(* IEC 61131-3 sources: daoli-st-library/DL_Process (part 11) *)

(* ---- FC_DL_CompressorDutyCycleCalc.st ---- *)
(*
  ============================================================
  组件名 : FC_DL_CompressorDutyCycleCalc
  分类   : DL_Process
  功能   : 压缩机加载占空比与卸载能耗占比计算，用于评估空压站运行经济性
  复杂度 : C1
  版本   : 1.0.0
  作者   : 道莅工业代码库工厂 / R81
  日期   : 2026-11-24
  开源溯源 : clean-room（no upstream）—— 依据公开工程公式自研，未复制任何上游实现
  红线自检 : R1 无GVL/R2 无物理地址/R3 纯IEC/R4 防除零/R5 双语注释
  接口说明 :
      加载占空比 = 加载时间 / 统计窗口 * 100。
      卸载能耗占比 = 卸载功率*卸载时间 / (加载功率*加载时间 + 卸载功率*卸载时间) * 100。
      能耗分母为零表示窗口内既无加载也无卸载，占空比无法归一，判无效。
      加载时间加卸载时间超过统计窗口时数据自相矛盾，判无效而不是强行归一。
  ============================================================
*)
FUNCTION FC_DL_CompressorDutyCycleCalc : BOOL
VAR_INPUT
    bEnable      : BOOL; // 使能：TRUE 时计算 / Enable: TRUE to compute
    bErr         : BOOL; // 外部故障：TRUE 时立即退出并置结果无效 / External fault: TRUE aborts with invalid result
    rLoadTime_s  : REAL; // 窗口内加载运行时间 [s] / loaded running time inside the window [second]
    rUnloadTime_s : REAL; // 窗口内卸载运行时间 [s] / unloaded running time inside the window [second]
    rIdleKw      : REAL; // 卸载空转功率 [kW] / unloaded idle power [kilowatt]
    rLoadKw      : REAL; // 加载运行功率 [kW] / loaded running power [kilowatt]
    rDur_s       : REAL; // 统计窗口总时长 [s] / total duration of the statistic window [second]
END_VAR
VAR_OUTPUT
    rDutyPct       : REAL; // 加载占空比，限幅 0~100 [%] / loading duty cycle clamped to 0 to 100 [percent]
    rIdleEnergyPct : REAL; // 卸载能耗占窗口总能耗比例，限幅 0~100 [%] / unloaded energy share of the window total clamped to 0 to 100 [percent]
    rTotalKwh      : REAL; // 窗口内折算总电量 [kWh] / equivalent total energy inside the window [kilowatt hour]
    bValid         : BOOL; // 输出有效：TRUE 表示结果可用 / Output valid
END_VAR
VAR CONSTANT
    DL_R_MAX   : REAL := 3.0E38;  // 实数上界，用于拦截 Inf [无量纲] / real upper bound used to reject infinity [dimensionless]
    DL_EPS     : REAL := 1.0E-12; // 除零判定阈值 [无量纲] / division guard threshold [dimensionless]
    DL_PCT     : REAL := 100.0;   // 百分数换算系数 [无量纲] / percentage scaling factor [dimensionless]
    DL_ZERO    : REAL := 0.0;     // 零值常量 [无量纲] / zero constant [dimensionless]
    DL_S_PER_H : REAL := 3600.0;  // 每小时秒数 [s/h] / seconds per hour [second per hour]
    DL_TOL_S   : REAL := 0.001;   // 时间窗超限判定容差 [s] / tolerance for the window overrun check [second]
END_VAR
VAR
    _bFin    : BOOL := FALSE; // 输入有限性判定结果 / input finiteness verdict
    _rLoadKwh : REAL := 0.0;  // 加载段电量 [kWh] / energy of the loaded segment [kilowatt hour]
    _rIdleKwh : REAL := 0.0;  // 卸载段电量 [kWh] / energy of the unloaded segment [kilowatt hour]
    _rDen     : REAL := 0.0;  // 能耗占比分母 [kWh] / denominator of the energy share [kilowatt hour]
END_VAR

    // 段 1｜出口预置
    rDutyPct := 0.0;
    rIdleEnergyPct := 0.0;
    rTotalKwh := 0.0;
    bValid := FALSE;
    // 段 2｜使能闸与外部故障闸
    IF NOT bEnable THEN
        RETURN;
    END_IF;
    IF bErr THEN
        RETURN;
    END_IF;
    // 段 3｜非有限闸
    _bFin := (rLoadTime_s = rLoadTime_s) AND (ABS(rLoadTime_s) <= DL_R_MAX) AND (rUnloadTime_s = rUnloadTime_s) AND (ABS(rUnloadTime_s) <= DL_R_MAX) AND (rIdleKw = rIdleKw) AND (ABS(rIdleKw) <= DL_R_MAX) AND (rLoadKw = rLoadKw) AND (ABS(rLoadKw) <= DL_R_MAX) AND (rDur_s = rDur_s) AND (ABS(rDur_s) <= DL_R_MAX);
    IF NOT _bFin THEN
        RETURN;
    END_IF;
    // 段 4｜域闸：统计窗口严格为正，时间与功率不得为负
    IF (ABS(rDur_s) <= DL_EPS) OR (rDur_s < DL_ZERO) THEN
        RETURN;
    END_IF;
    IF (rLoadTime_s < DL_ZERO) OR (rUnloadTime_s < DL_ZERO) OR (rIdleKw < DL_ZERO) OR (rLoadKw < DL_ZERO) THEN
        RETURN;
    END_IF;
    // 段 5｜加载加卸载不得超过窗口，超出部分属数据矛盾
    IF (rLoadTime_s + rUnloadTime_s) > (rDur_s + DL_TOL_S) THEN
        RETURN;
    END_IF;
    // 段 6｜加载占空比与限幅
    rDutyPct := rLoadTime_s / rDur_s * DL_PCT;
    IF rDutyPct < DL_ZERO THEN
        rDutyPct := DL_ZERO;
    END_IF;
    IF rDutyPct > DL_PCT THEN
        rDutyPct := DL_PCT;
    END_IF;
    // 段 7｜两段电量与总电量
    _rLoadKwh := rLoadKw * rLoadTime_s / DL_S_PER_H;
    _rIdleKwh := rIdleKw * rUnloadTime_s / DL_S_PER_H;
    rTotalKwh := _rLoadKwh + _rIdleKwh;
    // 段 8｜能耗占比分母闸
    _rDen := _rLoadKwh + _rIdleKwh;
    IF _rDen <= DL_EPS THEN
        RETURN;
    END_IF;
    rIdleEnergyPct := _rIdleKwh / _rDen * DL_PCT;
    IF rIdleEnergyPct < DL_ZERO THEN
        rIdleEnergyPct := DL_ZERO;
    END_IF;
    IF rIdleEnergyPct > DL_PCT THEN
        rIdleEnergyPct := DL_PCT;
    END_IF;
    bValid := TRUE;
    FC_DL_CompressorDutyCycleCalc := bValid;
END_FUNCTION

(* ---- FC_DL_ConductivityDilutionCalc.st ---- *)
(*
  ============================================================
  组件名 : FC_DL_ConductivityDilutionCalc
  分类   : DL_Process
  功能   : 电导率稀释比计算，由母液与水的本底电导求目标浓度所需的稀释倍数与配水占比
  复杂度 : C1
  版本   : 1.0.0
  作者   : 道莅工业代码库工厂 / R81
  日期   : 2026-11-24
  开源溯源 : clean-room（no upstream）—— 依据公开工程公式自研，未复制任何上游实现
  红线自检 : R1 无GVL/R2 无物理地址/R3 纯IEC/R4 防除零/R5 双语注释
  接口说明 :
      稀释比 = (母液电导 - 水本底电导) / (目标电导 - 水本底电导)。
      目标电导不高于水本底时分母非正，物理上无法靠兑水达到，直接判无效。
      配水占比 = (1 - 1/稀释比) * 100，稀释比非正时同样判无效。
  ============================================================
*)
FUNCTION FC_DL_ConductivityDilutionCalc : BOOL
VAR_INPUT
    bEnable      : BOOL; // 使能：TRUE 时计算 / Enable: TRUE to compute
    bErr         : BOOL; // 外部故障：TRUE 时立即退出并置结果无效 / External fault: TRUE aborts with invalid result
    rCondFeed    : REAL; // 母液电导率 [uS/cm] / feed solution conductivity [micro siemens per centimetre]
    rCondTarget  : REAL; // 目标电导率 [uS/cm] / target conductivity [micro siemens per centimetre]
    rCondWater   : REAL; // 稀释水本底电导率 [uS/cm] / background conductivity of the dilution water [micro siemens per centimetre]
END_VAR
VAR_OUTPUT
    rDilutionRatio : REAL; // 稀释倍数，母液体积的多少倍 [无量纲] / dilution ratio in multiples of the feed volume [dimensionless]
    rWaterPct      : REAL; // 配水中水所占体积百分比 [%] / volumetric percentage of water in the mixture [percent]
    bValid         : BOOL; // 输出有效：TRUE 表示结果可用 / Output valid
END_VAR
VAR CONSTANT
    DL_R_MAX : REAL := 3.0E38;  // 实数上界，用于拦截 Inf [无量纲] / real upper bound used to reject infinity [dimensionless]
    DL_EPS   : REAL := 1.0E-12; // 除零判定阈值 [无量纲] / division guard threshold [dimensionless]
    DL_ONE   : REAL := 1.0;     // 单位常量 [无量纲] / unity constant [dimensionless]
    DL_PCT   : REAL := 100.0;   // 百分数换算系数 [无量纲] / percentage scaling factor [dimensionless]
    DL_RATIO_MAX : REAL := 10000.0; // 稀释比合理上限，超限视为配比不可实现 [无量纲] / sanity upper bound of the dilution ratio [dimensionless]
END_VAR
VAR
    _bFin  : BOOL := FALSE; // 输入有限性判定结果 / input finiteness verdict
    _rNum  : REAL := 0.0;   // 稀释比分子 [uS/cm] / numerator of the dilution ratio [micro siemens per centimetre]
    _rDen  : REAL := 0.0;   // 稀释比分母 [uS/cm] / denominator of the dilution ratio [micro siemens per centimetre]
END_VAR

    // 段 1｜出口预置
    rDilutionRatio := 0.0;
    rWaterPct := 0.0;
    bValid := FALSE;
    // 段 2｜使能闸与外部故障闸
    IF NOT bEnable THEN
        RETURN;
    END_IF;
    IF bErr THEN
        RETURN;
    END_IF;
    // 段 3｜非有限闸
    _bFin := (rCondFeed = rCondFeed) AND (ABS(rCondFeed) <= DL_R_MAX) AND (rCondTarget = rCondTarget) AND (ABS(rCondTarget) <= DL_R_MAX) AND (rCondWater = rCondWater) AND (ABS(rCondWater) <= DL_R_MAX);
    IF NOT _bFin THEN
        RETURN;
    END_IF;
    // 段 4｜域闸：三者均不得为负，母液必须高于水本底
    IF (rCondFeed < 0.0) OR (rCondTarget < 0.0) OR (rCondWater < 0.0) THEN
        RETURN;
    END_IF;
    // 段 5｜分子分母组装
    _rNum := rCondFeed - rCondWater;
    _rDen := rCondTarget - rCondWater;
    // 段 6｜分母非正闸：兑水无法把电导降到水本底以下
    IF _rDen <= DL_EPS THEN
        RETURN;
    END_IF;
    // 段 7｜分子非正闸：母液不高于水本底时无稀释意义
    IF _rNum <= DL_EPS THEN
        RETURN;
    END_IF;
    rDilutionRatio := _rNum / _rDen;
    // 段 8｜稀释比合理区间闸，防止配比不可实现
    IF (rDilutionRatio < DL_ONE) OR (rDilutionRatio > DL_RATIO_MAX) THEN
        RETURN;
    END_IF;
    // 段 9｜配水占比
    rWaterPct := (DL_ONE - DL_ONE / rDilutionRatio) * DL_PCT;
    IF rWaterPct < 0.0 THEN
        rWaterPct := 0.0;
    END_IF;
    IF rWaterPct > DL_PCT THEN
        rWaterPct := DL_PCT;
    END_IF;
    bValid := TRUE;
    FC_DL_ConductivityDilutionCalc := bValid;
END_FUNCTION

(* ---- FC_DL_CoreSandBakeCurveCalc.st ---- *)
(*
 * FC_DL_CoreSandBakeCurveCalc | C2 | DL_Process
 * 功能：芯砂烘干升温曲线（升温段、总时间）与保温后残余水分       单位：温度 [℃]、升温速率 [K/min]、时间 [min]、水分 [%]
 * 工况边界：升温段按线性斜坡、保温段按一阶指数衰减残余水分 res=1.5×EXP(−hold/40)；升温速率须 >0、目标温度须高于起始温度，否则判 9716；本件不含分段升温与露点控制
 * 代数值回代：target=200、start=25、rate=3 → ramp=175/3=58.33 min；total=58.33+60=118.33 min；res=1.5×EXP(−60/40)=1.5×0.2231=0.335 %（spec 记 0.33 %，一致）
 * 开源溯源：clean-room 自研，未复制任何第三方代码（无外部来源）
 *)
FUNCTION FC_DL_CoreSandBakeCurveCalc : BOOL
VAR_INPUT
    rTargetC   : REAL := 200.0;      // 目标烘干温度 | target baking temperature [℃]
    rRampKmin  : REAL := 3.0;        // 升温速率 | heating rate [K/min]
    rStartC    : REAL := 25.0;       // 起始温度 | starting temperature [℃]
    rHoldMin   : REAL := 60.0;       // 保温时间 | holding time [min]
END_VAR
VAR_OUTPUT
    rRampMin        : REAL;          // 升温段时间 | ramp duration [min]
    rTotalMin       : REAL;          // 总时间（升温+保温）| total time, ramp plus hold [min]
    rResidualMoistPct : REAL;        // 保温后残余水分 | residual moisture after holding [%]
    xValid          : BOOL;          // 输出有效 | outputs valid
    nFaultCode      : INT;           // 0=无 / 9716=温度或速率非法 | 0 none, 9716 illegal temperature or rate
END_VAR
VAR
    xFinTg  : BOOL;                  // 目标温度有限性 | target temperature is finite
    xFinRt  : BOOL;                  // 升温速率有限性 | heating rate is finite
    xFinSt  : BOOL;                  // 起始温度有限性 | starting temperature is finite
    xFinHd  : BOOL;                  // 保温时间有限性 | holding time is finite
END_VAR
VAR CONSTANT
    DL_CSB_MOIST0   : REAL := 1.5;   // 保温起始残余水分基准 | residual moisture at the start of holding [%]
    DL_CSB_TAU_MIN  : REAL := 40.0;  // 水分衰减时间常数 | moisture decay time constant [min]
END_VAR

// 段1｜非有限闸（R19）
xFinTg := (rTargetC = rTargetC) AND ((rTargetC - rTargetC) = 0.0);
xFinRt := (rRampKmin = rRampKmin) AND ((rRampKmin - rRampKmin) = 0.0);
xFinSt := (rStartC = rStartC) AND ((rStartC - rStartC) = 0.0);
xFinHd := (rHoldMin = rHoldMin) AND ((rHoldMin - rHoldMin) = 0.0);
IF (NOT xFinTg) OR (NOT xFinRt) OR (NOT xFinSt) OR (NOT xFinHd) THEN
    rRampMin := 0.0;                 // 安全值：时间 0 | safe value, zero times
    rTotalMin := 0.0;
    rResidualMoistPct := 0.0;
    xValid := FALSE;
    nFaultCode := 9716;
    FC_DL_CoreSandBakeCurveCalc := FALSE;
    RETURN;
END_IF

// 段2｜域闸：速率入分母须 >0，目标须高于起始，保温时间非负
IF (rRampKmin <= 0.0) OR (rTargetC <= rStartC) OR (rHoldMin < 0.0) THEN
    rRampMin := 0.0;
    rTotalMin := 0.0;
    rResidualMoistPct := 0.0;
    xValid := FALSE;
    nFaultCode := 9716;
    FC_DL_CoreSandBakeCurveCalc := FALSE;
    RETURN;
END_IF

// 段3｜算法：ramp=(target−start)/rate；total=ramp+hold；res=1.5×EXP(−hold/40)
rRampMin := (rTargetC - rStartC) / rRampKmin;
rTotalMin := rRampMin + rHoldMin;
rResidualMoistPct := DL_CSB_MOIST0 * EXP(-rHoldMin / DL_CSB_TAU_MIN);

// 段4｜出口
nFaultCode := 0;
xValid := TRUE;
FC_DL_CoreSandBakeCurveCalc := TRUE;
END_FUNCTION

(* ---- FC_DL_CrusherThroughputCalc.st ---- *)
(*
  Name: FC_DL_CrusherThroughputCalc
  Category: DL_Process
  Version: 1.0.0
  Round: R89 / 2026-11-25
  开源溯源：clean-room 自研（族 矿山破碎筛分，ST 开源生态实测 0 命中，无外部代码引入）
  功能：按排矿口开口比产能法算颚式/圆锥破碎机实际产能，并以单程合格率反算闭路循环负荷率。
  边界条件：① 五入参全部过非有限闸（NaN 自反判 / Inf 差值自减判），任一非有限返回哨兵 -1；
            ② 排矿口 < 3 mm 或给料粒度不高于排矿口 1.2 倍（无有效破碎比）判组态非法，返回哨兵 -1；
            ③ 单程合格率下限 0.1，循环负荷率钳位 0~500 %（钳的是量值不钳事实，有效性不受影响）。
  量纲自证：q0[t/(h·mm)] × gap[mm] = t/h；kH / kD 无量纲；CL=(1/p−1)×100 无量纲。
*)
FUNCTION FC_DL_CrusherThroughputCalc : REAL
VAR_INPUT
    fFeedTph : REAL;        (* 给料量（新给矿） [t/h] Feed rate, fresh feed *)
    fGapMm : REAL;          (* 排矿口开口（闭侧） [mm] Closed-side gap [mm] *)
    fFeedSizeMm : REAL;     (* 给料粒度（95% 通过粒径） [mm] Feed size, 95% passing *)
    fHardnessIdx : REAL;    (* 硬度指数（1.0 为基准矿） [-] Hardness index, 1.0 baseline *)
    fBulkDensity : REAL;    (* 堆密度 [t/m3] Bulk density [t/m3] *)
END_VAR
VAR_OUTPUT
    fThroughputTph : REAL;      (* 实际破碎通过量 [t/h] Actual throughput [t/h] *)
    fCirculatingLoadPct : REAL; (* 闭路循环负荷率 [%] Circulating load ratio [%] *)
    xValid : BOOL;              (* 计算有效性标志 [-] Calculation valid flag *)
END_VAR
VAR CONSTANT
    DL_EPS : REAL := 1.0E-9;        (* 除零判定容差 [-] Divide-by-zero tolerance *)
    DL_Q0 : REAL := 2.5;            (* 单位开口基准产能 [t/(h·mm)] Specific capacity per gap *)
    DL_DENS_REF : REAL := 1.6;      (* 基准堆密度 [t/m3] Reference bulk density *)
    DL_RR_MIN : REAL := 1.2;        (* 最小有效破碎比 [-] Minimum reduction ratio *)
    DL_CL_MAX : REAL := 500.0;      (* 循环负荷率饱和上限 [%] Circulating load ceiling *)
    DL_PASS_MIN : REAL := 0.1;      (* 单程合格率下限 [-] Minimum single-pass fraction *)
    DL_GAP_MIN : REAL := 3.0;       (* 排矿口工程下限 [mm] Minimum engineering gap *)
    DL_H_MIN : REAL := 0.2;         (* 硬度指数下限 [-] Hardness index floor *)
    DL_H_MAX : REAL := 5.0;         (* 硬度指数上限 [-] Hardness index ceiling *)
    DL_D_MIN : REAL := 0.5;         (* 堆密度下限 [t/m3] Bulk density floor *)
    DL_D_MAX : REAL := 4.0;         (* 堆密度上限 [t/m3] Bulk density ceiling *)
END_VAR
VAR
    fRr : REAL;     (* 破碎比 = 给料粒度/排矿口 [-] Reduction ratio *)
    fKh : REAL;     (* 硬度修正系数 [-] Hardness correction factor *)
    fKd : REAL;     (* 密度修正系数 [-] Density correction factor *)
    fQcap : REAL;   (* 排矿口通过能力 [t/h] Gap capability [t/h] *)
    fPass : REAL;   (* 单程合格率 [-] Single-pass pass fraction *)
    fQout : REAL;   (* 当拍通过量中间量 [t/h] Throughput scratch [t/h] *)
END_VAR
(* 出口预置：三出口统一预置安全值（R256） *)
fThroughputTph := 0.0; fCirculatingLoadPct := 0.0; xValid := FALSE;
(* 非有限闸：NaN 自反判 + Inf 差值自减判，五入参全枚举（R272） *)
IF (fFeedTph <> fFeedTph) OR ((fFeedTph - fFeedTph) <> 0.0)
   OR (fGapMm <> fGapMm) OR ((fGapMm - fGapMm) <> 0.0)
   OR (fFeedSizeMm <> fFeedSizeMm) OR ((fFeedSizeMm - fFeedSizeMm) <> 0.0)
   OR (fHardnessIdx <> fHardnessIdx) OR ((fHardnessIdx - fHardnessIdx) <> 0.0)
   OR (fBulkDensity <> fBulkDensity) OR ((fBulkDensity - fBulkDensity) <> 0.0) THEN
    FC_DL_CrusherThroughputCalc := -1.0;    (* 哨兵 -1：入参非有限 / Sentinel -1, non-finite input *)
    RETURN;
END_IF
(* 组态域闸：给料、开口、粒度、硬度、密度逐项定域（禁 NaN 判假即放行，全用正向不等号） *)
IF (fFeedTph <= DL_EPS) OR (fGapMm < DL_GAP_MIN)
   OR (fFeedSizeMm <= fGapMm * DL_RR_MIN)
   OR (fHardnessIdx < DL_H_MIN) OR (fHardnessIdx > DL_H_MAX)
   OR (fBulkDensity < DL_D_MIN) OR (fBulkDensity > DL_D_MAX) THEN
    FC_DL_CrusherThroughputCalc := -1.0;    (* 哨兵 -1：组态非法 / Sentinel -1, bad configuration *)
    RETURN;
END_IF
(* 破碎比：给料粒度 ÷ 排矿口，除子已过工程下限闸，量纲 mm/mm = 无量纲 *)
fRr := fFeedSizeMm / fGapMm;
(* 硬度修正：kH = 1/(0.6+0.4·H)，H = 1.0 时恰为 1.0，硬矿按比例降产能 *)
fKh := 1.0 / (0.6 + 0.4 * fHardnessIdx);
(* 密度修正：kD = ρ/ρref，无量纲 *)
fKd := fBulkDensity / DL_DENS_REF;
(* 排矿口通过能力：q0[t/(h·mm)] × gap[mm] × kH × kD，量纲收敛为 t/h *)
fQcap := DL_Q0 * fGapMm * fKh * fKd;
(* 实际通过量取给料与能力较小者：能力不足即积料，不虚报产能 *)
IF fFeedTph > fQcap THEN
    fQout := fQcap;
ELSE
    fQout := fFeedTph;
END_IF
(* 单程合格率：p = 1/(1+0.5·(Rr−1))，破碎比越大单程越粗、合格率越低 *)
fPass := 1.0 / (1.0 + 0.5 * (fRr - 1.0));
IF fPass < DL_PASS_MIN THEN
    fPass := DL_PASS_MIN;                   (* 下限钳位，防循环负荷率发散 / Clamp to avoid divergence *)
END_IF
(* 循环负荷率：CL = (1/p − 1)×100，除子 p 已过下限钳位，绝无零除 *)
fThroughputTph := fQout;
fCirculatingLoadPct := (1.0 / fPass - 1.0) * 100.0;
IF fCirculatingLoadPct > DL_CL_MAX THEN
    fCirculatingLoadPct := DL_CL_MAX;       (* 量值饱和钳位（事实量不饱和） / Value saturation *)
END_IF
xValid := TRUE;                             (* 链路有效 / Chain valid *)
FC_DL_CrusherThroughputCalc := fThroughputTph;
END_FUNCTION

(* ---- FC_DL_CutLengthDeviationCalc.st ---- *)
(*
  DL Factory R83 | FC_DL_CutLengthDeviationCalc
  功能：比较定长裁切设定值与实测值，输出偏差、反向补偿量并做死区判稳。
  开源溯源：无（clean-room 自研，依据公开工艺公式，来源=行业通用公式，许可证=MIT，借鉴点=公式结构）
  规则：R1-R21 全遵守
*)
FUNCTION FC_DL_CutLengthDeviationCalc : REAL
VAR_INPUT
    fSetLenMm   : REAL; // 定长设定值 [mm] / Cut length setpoint [mm]
    fMeasLenMm  : REAL; // 实测裁切长度 [mm] / Measured cut length [mm]
    fDeadbandMm : REAL; // 死区（不补偿带宽）[mm] / Deadband, no-compensation band [mm]
    fCompGain   : REAL; // 补偿增益（0~200）[%] / Compensation gain [%]
END_VAR
VAR_OUTPUT
    fDevMm  : REAL; // 长度偏差（实测-设定，正=偏长）[mm] / Deviation, + = too long [mm]
    fCompMm : REAL; // 补偿量（叠加设定值，符号与偏差相反）[mm] / Compensation to add [mm]
    xInBand : BOOL; // 在死区内（TRUE=无需补偿）/ Inside deadband, TRUE = no trim
END_VAR
VAR
    fAbsDev : REAL; // 偏差绝对值 [mm] / Absolute deviation [mm]
    fGainK  : REAL; // 增益归一化系数 [-]/ Normalised gain factor
END_VAR
// 出口预置：预置在带内（无动作安全侧），非有限拍不产生补偿
fDevMm := 0.0; fCompMm := 0.0; xInBand := TRUE;
// 非有限拦截 + 量纲自检（R20/R21）
IF NOT (fSetLenMm > -1.0E30 AND fSetLenMm < 1.0E30) OR NOT (fMeasLenMm > -1.0E30 AND fMeasLenMm < 1.0E30) OR NOT (fDeadbandMm > -1.0E30 AND fDeadbandMm < 1.0E30) OR NOT (fCompGain > -1.0E30 AND fCompGain < 1.0E30) OR fSetLenMm <= 0.0 OR fDeadbandMm < 0.0 THEN
    FC_DL_CutLengthDeviationCalc := -1.0; RETURN;  // 哨兵 -1：非有限或量纲越界 / Sentinel -1
END_IF
// 增益域闸：0~200% 之外按边界钳位后继续
IF fCompGain < 0.0 THEN
    fGainK := 0.0;                  // 负增益等价不补偿 [-] / Negative gain equals no compensation
ELSIF fCompGain > 200.0 THEN
    fGainK := 2.0;                  // 增益上限 2.0 倍 [-] / Gain clamped to 2.0
ELSE
    fGainK := fCompGain / 100.0;    // 归一化增益 [-] / Normalised gain
END_IF
// 偏差：实测减设定，同量纲（mm）直接相减
fDevMm  := fMeasLenMm - fSetLenMm;   // 长度偏差 [mm] / Length deviation [mm]
fAbsDev := ABS(fDevMm);              // 偏差绝对值 [mm] / Absolute deviation [mm]
// 死区判定与补偿：带内不补偿，带外按增益反向补偿（浮点比较只用绝对差与不等）
IF fAbsDev <= fDeadbandMm THEN
    xInBand := TRUE;                 // 在死区内不动作 / In deadband, no action
    fCompMm := 0.0;                  // 补偿量为零 [mm] / Compensation zero
ELSE
    xInBand := FALSE;                // 越出死区 / Outside deadband
    fCompMm := -fDevMm * fGainK;     // 反向补偿量 [mm] / Reverse compensation [mm]
END_IF
FC_DL_CutLengthDeviationCalc := fDevMm;   // 返回长度偏差 [mm] / Return deviation [mm]
END_FUNCTION

(* ---- FC_DL_CutTobaccoFinesCalc.st ---- *)
(*
 * FC_DL_CutTobaccoFinesCalc | C1 | DL_Process
 * 功能：碎丝率（≤0.5 mm 占比）与整丝率（≥2.5 mm 占比）       单位：质量 [g]、占比 [%]
 * 工况边界：样品质量须 >0（入分母）；两率之和 >100 % 说明筛分数据自相矛盾，判 9511；筛网规格固定为 0.5 mm 与 2.5 mm，更换筛网须重新标定；中间档丝（0.5~2.5 mm）占比作为信息量输出
 * 代数值回代：m=100 g、fines=8 g、long=85 g → 碎丝率 8.0 %、整丝率 85.0 %、中间档 7.0 %（合计 100 %，与 spec 判定式一致）
 * 开源溯源：clean-room 自研，未复制任何第三方代码（无外部来源）
 *)
FUNCTION FC_DL_CutTobaccoFinesCalc : BOOL
VAR_INPUT
    rSampleG : REAL := 100.0;        // 样品总质量 | total sample mass [g]
    rFinesG  : REAL;                 // 碎丝质量（≤0.5 mm）| fines mass, 0.5 mm and below [g]
    rLongG   : REAL;                 // 整丝质量（≥2.5 mm）| long strands, 2.5 mm and above [g]
END_VAR
VAR_OUTPUT
    rFinesPct : REAL;                // 碎丝率 | fines ratio [%]
    rLongPct  : REAL;                // 整丝率 | long strand ratio [%]
    rMidPct   : REAL;                // 中间档占比（信息量）| middle fraction ratio, informational [%]
    xValid    : BOOL;                // 输出有效 | outputs valid
    nFaultCode: INT;                 // 0=无 / 9511=样品或筛分数据非法 | 0 none, 9511 illegal sample or sieve data
END_VAR
VAR
    xFinS : BOOL;                    // 样品质量有限性 | sample mass is finite
    xFinF : BOOL;                    // 碎丝质量有限性 | fines mass is finite
    xFinL : BOOL;                    // 整丝质量有限性 | long strand mass is finite
    rSumPct : REAL;                  // 两率之和 | sum of the two ratios [%]
END_VAR
VAR CONSTANT
    DL_CTF_PCT     : REAL := 100.0;  // 百分数换算系数 | percentage factor [%]
    DL_CTF_S_MIN   : REAL := 1.0E-6; // 样品质量下限（防零除）| sample mass lower bound [g]
    DL_CTF_SUM_MAX : REAL := 100.0;  // 两率之和上限 | upper bound of the summed ratios [%]
    DL_CTF_EPS     : REAL := 1.0E-6; // 浮点比较容差 | floating comparison tolerance [%]
END_VAR

// 段1｜非有限闸（R19）
xFinS := (rSampleG = rSampleG) AND ((rSampleG - rSampleG) = 0.0);
xFinF := (rFinesG = rFinesG) AND ((rFinesG - rFinesG) = 0.0);
xFinL := (rLongG = rLongG) AND ((rLongG - rLongG) = 0.0);
IF (NOT xFinS) OR (NOT xFinF) OR (NOT xFinL) THEN
    rFinesPct := 0.0;                // 安全值：两率 0 | safe value, zero ratios
    rLongPct := 0.0;
    rMidPct := 0.0;
    xValid := FALSE;
    nFaultCode := 9511;
    FC_DL_CutTobaccoFinesCalc := FALSE;
    RETURN;
END_IF

// 段2｜域闸：样品质量入分母必须 >0，两档质量不得为负
IF (rSampleG <= DL_CTF_S_MIN) OR (rFinesG < 0.0) OR (rLongG < 0.0) THEN
    rFinesPct := 0.0;
    rLongPct := 0.0;
    rMidPct := 0.0;
    xValid := FALSE;
    nFaultCode := 9511;
    FC_DL_CutTobaccoFinesCalc := FALSE;
    RETURN;
END_IF

// 段3｜算法：两率各按样品总量计算
rFinesPct := rFinesG / rSampleG * DL_CTF_PCT;
rLongPct := rLongG / rSampleG * DL_CTF_PCT;
rSumPct := rFinesPct + rLongPct;

// 段4｜数据自洽校验：两率之和不得超过 100 %
IF rSumPct > (DL_CTF_SUM_MAX + DL_CTF_EPS) THEN
    rMidPct := 0.0;                  // 安全值：中间档置 0 | safe value, middle fraction zeroed
    xValid := FALSE;
    nFaultCode := 9511;
    FC_DL_CutTobaccoFinesCalc := FALSE;
    RETURN;
END_IF

// 段5｜中间档与出口
rMidPct := DL_CTF_SUM_MAX - rSumPct;
nFaultCode := 0;
xValid := TRUE;
FC_DL_CutTobaccoFinesCalc := TRUE;
END_FUNCTION

(* ---- FC_DL_CutTobaccoWidthCalc.st ---- *)
(*
 * FC_DL_CutTobaccoWidthCalc | C2 | DL_Process
 * 功能：由线速、刀辊转速与刀片数推算切丝宽度并判定丝宽合格       单位：线速 [m/s]、转速 [r/min]、刀数 [片]、丝宽 [mm]
 * 工况边界：nRpm 与 nBlades 须 >0（入分母），线速须 ≥0 且有限；仅适用于定刀数圆盘切丝机，不含刀片磨损补偿；入参非法一律 xValid=FALSE 且丝宽取 0
 * 代数值回代：v=0.5 m/s、rpm=3000、blades=10 → w=0.5×1000×60/(3000×10)=1.0 mm，目标 1.0 mm → 合格（与 spec 回代行一致）
 * 开源溯源：clean-room 自研，未复制任何第三方代码（无外部来源）
 *)
FUNCTION FC_DL_CutTobaccoWidthCalc : BOOL
VAR_INPUT
    rLineSpeedMps : REAL;            // 烟片线速度 | tobacco line speed [m/s]
    nRpm          : INT;             // 刀辊转速 | cutter drum speed [r/min]
    nBlades       : INT;             // 刀片数 | blade count [片]
    rTargetMm     : REAL := 1.0;     // 目标丝宽 | target cut width [mm]
    rTolMm        : REAL := 0.1;     // 丝宽公差（±）| cut width tolerance [mm]
END_VAR
VAR_OUTPUT
    rWidthMm      : REAL;            // 实际丝宽 | actual cut width [mm]
    rDevMm        : REAL;            // 相对目标的偏差 | deviation from the target [mm]
    xInTolerance  : BOOL;            // 丝宽在公差带内 | cut width within tolerance
    xValid        : BOOL;            // 输出有效 | outputs valid
END_VAR
VAR
    xFinV  : BOOL;                   // 线速有限性 | line speed is finite
    xFinTg : BOOL;                   // 目标有限性 | target is finite
    xFinTol: BOOL;                   // 公差有限性 | tolerance is finite
    rRpm   : REAL;                   // 转速的实数形式 | drum speed as a real number [r/min]
    rBlades: REAL;                   // 刀数的实数形式 | blade count as a real number [片]
    rDen   : REAL;                   // 分母（转速×刀数）| denominator, speed times blade count [1/min]
END_VAR
VAR CONSTANT
    DL_CTW_SEC_PER_MIN : REAL := 60.0;      // 分转秒系数 | minutes to seconds factor [s/min]
    DL_CTW_M_TO_MM     : REAL := 1000.0;    // 米转毫米系数 | metres to millimetres factor [mm/m]
    DL_CTW_DEN_MIN     : REAL := 1.0E-9;    // 除零保护阈值 | division guard threshold [1/min]
    DL_CTW_TOL_EPS     : REAL := 1.0E-6;    // 浮点比较容差 | floating comparison tolerance [mm]
END_VAR

// 段1｜非有限闸（R19）
xFinV := (rLineSpeedMps = rLineSpeedMps) AND ((rLineSpeedMps - rLineSpeedMps) = 0.0);
xFinTg := (rTargetMm = rTargetMm) AND ((rTargetMm - rTargetMm) = 0.0);
xFinTol := (rTolMm = rTolMm) AND ((rTolMm - rTolMm) = 0.0);
IF (NOT xFinV) OR (NOT xFinTg) OR (NOT xFinTol) THEN
    rWidthMm := 0.0;                 // 安全值：丝宽 0 | safe value, zero width
    rDevMm := 0.0;
    xInTolerance := FALSE;
    xValid := FALSE;
    FC_DL_CutTobaccoWidthCalc := FALSE;
    RETURN;
END_IF

// 段2｜域闸：转速与刀数必须为正（入分母），线速不得为负，公差须为正
IF (nRpm <= 0) OR (nBlades <= 0) OR (rLineSpeedMps < 0.0) OR (rTolMm <= 0.0) THEN
    rWidthMm := 0.0;
    rDevMm := 0.0;
    xInTolerance := FALSE;
    xValid := FALSE;
    FC_DL_CutTobaccoWidthCalc := FALSE;
    RETURN;
END_IF

// 段3｜算法：w_mm = (v×1000×60)/(rpm×nBlades)，分母显式防零
rRpm := INT_TO_REAL(nRpm);
rBlades := INT_TO_REAL(nBlades);
rDen := rRpm * rBlades;
IF rDen > DL_CTW_DEN_MIN THEN
    rWidthMm := (rLineSpeedMps * DL_CTW_M_TO_MM * DL_CTW_SEC_PER_MIN) / rDen;
ELSE
    rWidthMm := 0.0;                 // 理论不可达（段2已排除），防御性兜底 | unreachable defence
END_IF

// 段4｜合格判定：偏差与公差同源于原始丝宽（R24）
rDevMm := rWidthMm - rTargetMm;
xInTolerance := ABS(rDevMm) <= (rTolMm + DL_CTW_TOL_EPS);
xValid := TRUE;
FC_DL_CutTobaccoWidthCalc := TRUE;
END_FUNCTION

(* ---- FC_DL_DemisterVelocityChk.st ---- *)
(*
  道莅工业代码库 / Daoli Industrial ST Library
  组件: FC_DL_DemisterVelocityChk
  分类: DL_Process
  开源溯源: 无（clean-room 工程公式自研；参考公开工艺计算公式，未复制任何受版权保护代码）
  许可证: 本项目自有 (MIT)
  功能: 除雾器截面气速与临界携带速度（Souders-Brown）比较，判定雾沫夹带
*)
FUNCTION FC_DL_DemisterVelocityChk : BOOL
VAR_INPUT
    rGasM3h : REAL; // 实际工况烟气量 [m3/h] / actual gas flow
    rAreaM2 : REAL; // 除雾器有效流通面积 [m2] / demister free area
    rRhoL : REAL; // 液相密度 [kg/m3] / liquid density
    rRhoG : REAL; // 气相密度 [kg/m3] / gas density
    rKFactor : REAL; // Souders-Brown 经验系数 [m/s] / Souders-Brown coefficient
END_VAR
VAR_OUTPUT
    rVelMs : REAL; // 截面气速 [m/s] / superficial gas velocity
    rVcritMs : REAL; // 临界夹带速度 [m/s] / critical carry-over velocity
    bValid : BOOL; // 结果有效位 [-] / result valid flag
    bCarryOver : BOOL; // 雾沫夹带标志（气速超临界）[-] / carry-over flag
    iErrCode : INT; // 事件码 0=正常 1=气相密度非法 2=流通面积非法 3=密度差不正 4=结果非有限 / event code
END_VAR
VAR CONSTANT
    rSecPerHour : REAL := 3600.0; // 每小时秒数 [s/h] / seconds per hour
END_VAR
VAR
    rRhoRatio : REAL; // 密度比 (ρL-ρG)/ρG [-] / density ratio
    rVelRaw : REAL; // 未限幅气速 [m/s] / unlimited velocity
    rVcritRaw : REAL; // 未限幅临界速度 [m/s] / unlimited critical velocity
END_VAR

    // —— 段 0：全路径预清 —— //
    rRhoRatio := 0.0;
    rVelRaw := 0.0;
    rVcritRaw := 0.0;
    rVelMs := 0.0;
    rVcritMs := 0.0;
    bValid := FALSE;
    bCarryOver := FALSE;
    iErrCode := 0;
    FC_DL_DemisterVelocityChk := FALSE;
    // —— 段 1：分母闸（气相密度、流通面积） —— //
    IF rRhoG <= 0.0 THEN
        iErrCode := 1; // 气相密度非法，临界速度无定义 / invalid gas density
        RETURN;
    END_IF;
    IF rAreaM2 <= 0.0 THEN
        iErrCode := 2; // 流通面积非法，气速无定义 / invalid free area
        RETURN;
    END_IF;
    // —— 段 2：截面气速（量纲 (m3/h)/(s/h)/(m2) = m/s） —— //
    rVelRaw := rGasM3h / rSecPerHour / rAreaM2; // 截面气速 [m/s] / superficial velocity
    IF ABS(rVelRaw) > 1.0E15 THEN
        iErrCode := 4; // 结果非有限，强制归零 / non-finite result, forced to zero
        RETURN;
    END_IF;
    IF rVelRaw < 0.0 THEN
        rVelMs := 0.0; // 负流量防御 / negative flow guard
    ELSE
        rVelMs := rVelRaw;
    END_IF;
    // —— 段 3：临界速度 = K·SQRT((ρL-ρG)/ρG)（开方前闸 >= 0） —— //
    rRhoRatio := (rRhoL - rRhoG) / rRhoG; // 密度比 [-] / density ratio
    IF rRhoRatio < 0.0 THEN
        rVcritMs := 0.0;
        iErrCode := 3; // 密度差不正（气相重于液相），临界速度无意义 / non-positive density difference
        bValid := TRUE;
        FC_DL_DemisterVelocityChk := TRUE;
        RETURN;
    END_IF;
    rVcritRaw := rKFactor * SQRT(rRhoRatio); // 临界速度 [m/s] / critical velocity
    IF ABS(rVcritRaw) > 1.0E15 THEN
        rVcritMs := 0.0;
        iErrCode := 4; // 结果非有限，强制归零 / non-finite result, forced to zero
        RETURN;
    END_IF;
    IF rVcritRaw < 0.0 THEN
        rVcritMs := 0.0; // 负系数防御 / negative coefficient guard
    ELSE
        rVcritMs := rVcritRaw;
    END_IF;
    // —— 段 4：夹带判定与收口 —— //
    bCarryOver := rVelMs > rVcritMs; // 夹带标志 [-] / carry-over flag
    bValid := TRUE;
    FC_DL_DemisterVelocityChk := TRUE;
END_FUNCTION

(* ---- FC_DL_DesiccantLifeEstimate.st ---- *)
(*
  ============================================================
  组件名 : FC_DL_DesiccantLifeEstimate
  分类   : DL_Process
  功能   : 干燥剂寿命估算，按累计吸湿量与温度降额后的有效容量求剩余寿命百分比
  复杂度 : C1
  版本   : 1.0.0
  作者   : 道莅工业代码库工厂 / R81
  日期   : 2026-11-24
  开源溯源 : clean-room（no upstream）—— 依据公开工程公式自研，未复制任何上游实现
  红线自检 : R1 无GVL/R2 无物理地址/R3 纯IEC/R4 防除零/R5 双语注释
  接口说明 :
      有效容量 = 额定吸附容量 * 温度降额系数，温度降额系数限定 0~1 区间且必须为正。
      剩余百分比 = (1 - 累计吸湿量/有效容量) * 100，限幅 0~100。
      剩余低于 20% 判更换到期；累计吸湿量超过有效容量时剩余按 0 截断，判定仍成立。
  ============================================================
*)
FUNCTION FC_DL_DesiccantLifeEstimate : BOOL
VAR_INPUT
    bEnable        : BOOL; // 使能：TRUE 时估算 / Enable: TRUE to estimate
    bErr           : BOOL; // 外部故障：TRUE 时立即退出并置结果无效 / External fault: TRUE aborts with invalid result
    rMoistureLoad  : REAL; // 累计已吸附水汽质量 [g] / accumulated adsorbed moisture mass [gram]
    rCapG          : REAL; // 额定吸附容量 [g] / rated adsorption capacity [gram]
    rTempDerate    : REAL; // 温度降额系数，1 表示不降额 [无量纲] / temperature derating factor, one means no derating [dimensionless]
END_VAR
VAR_OUTPUT
    rEffCapG   : REAL; // 降额后的有效吸附容量 [g] / effective capacity after derating [gram]
    rLoadPct   : REAL; // 已消耗容量百分比 [%] / consumed capacity percentage [percent]
    rRemainPct : REAL; // 剩余寿命百分比，限幅 0~100 [%] / remaining life percentage clamped to 0 to 100 [percent]
    bReplaceDue : BOOL; // 更换到期：TRUE 表示剩余低于 20% / replacement due, TRUE when the remainder is below 20 percent
    bValid     : BOOL; // 输出有效：TRUE 表示结果可用 / Output valid
END_VAR
VAR CONSTANT
    DL_R_MAX   : REAL := 3.0E38; // 实数上界，用于拦截 Inf [无量纲] / real upper bound used to reject infinity [dimensionless]
    DL_EPS     : REAL := 1.0E-12; // 除零判定阈值 [无量纲] / division guard threshold [dimensionless]
    DL_ONE     : REAL := 1.0;     // 单位常量 [无量纲] / unity constant [dimensionless]
    DL_ZERO    : REAL := 0.0;     // 零值常量 [无量纲] / zero constant [dimensionless]
    DL_PCT     : REAL := 100.0;   // 百分数换算系数 [无量纲] / percentage scaling factor [dimensionless]
    DL_DUE_PCT : REAL := 20.0;    // 更换到期门限 [%] / replacement due threshold [percent]
END_VAR
VAR
    _bFin : BOOL := FALSE; // 输入有限性判定结果 / input finiteness verdict
    _rUse : REAL := 0.0;   // 容量占用比 [无量纲] / capacity usage ratio [dimensionless]
END_VAR

    // 段 1｜出口预置：剩余先置 0（最不利），防止下游误判为充足
    rEffCapG := 0.0;
    rLoadPct := 0.0;
    rRemainPct := 0.0;
    bReplaceDue := TRUE;
    bValid := FALSE;
    // 段 2｜使能闸与外部故障闸
    IF NOT bEnable THEN
        RETURN;
    END_IF;
    IF bErr THEN
        RETURN;
    END_IF;
    // 段 3｜非有限闸
    _bFin := (rMoistureLoad = rMoistureLoad) AND (ABS(rMoistureLoad) <= DL_R_MAX) AND (rCapG = rCapG) AND (ABS(rCapG) <= DL_R_MAX) AND (rTempDerate = rTempDerate) AND (ABS(rTempDerate) <= DL_R_MAX);
    IF NOT _bFin THEN
        RETURN;
    END_IF;
    // 段 4｜域闸：容量严格为正，降额系数落在 0~1 且严格为正
    IF (ABS(rCapG) <= DL_EPS) OR (rCapG < DL_ZERO) THEN
        RETURN;
    END_IF;
    IF (ABS(rTempDerate) <= DL_EPS) OR (rTempDerate < DL_ZERO) OR (rTempDerate > DL_ONE) THEN
        RETURN;
    END_IF;
    IF rMoistureLoad < DL_ZERO THEN
        RETURN;
    END_IF;
    // 段 5｜有效容量：容量乘降额系数，乘积仍须严格为正才可作分母
    rEffCapG := rCapG * rTempDerate;
    IF rEffCapG <= DL_EPS THEN
        RETURN;
    END_IF;
    // 段 6｜占用比与剩余百分比
    _rUse := rMoistureLoad / rEffCapG;
    rLoadPct := _rUse * DL_PCT;
    rRemainPct := (DL_ONE - _rUse) * DL_PCT;
    // 段 7｜限幅
    IF rRemainPct < DL_ZERO THEN
        rRemainPct := DL_ZERO;
    END_IF;
    IF rRemainPct > DL_PCT THEN
        rRemainPct := DL_PCT;
    END_IF;
    IF rLoadPct < DL_ZERO THEN
        rLoadPct := DL_ZERO;
    END_IF;
    // 段 8｜更换到期判定
    IF rRemainPct < DL_DUE_PCT THEN
        bReplaceDue := TRUE;
    ELSE
        bReplaceDue := FALSE;
    END_IF;
    bValid := TRUE;
    FC_DL_DesiccantLifeEstimate := bValid;
END_FUNCTION

(* ---- FC_DL_DewaterMassBalance.st ---- *)
(*
  道莅工业代码库 / Daoli Industrial ST Library
  组件: FC_DL_DewaterMassBalance
  分类: DL_Process
  开源溯源: 无（clean-room 工程公式自研；参考公开工艺计算公式，未复制任何受版权保护代码）
  许可证: 本项目自有 (MIT)
  功能: 脱水单元干固体质量平衡：由进泥与泥饼含固率反算泥饼量、滤液量与固体回收率
*)
FUNCTION FC_DL_DewaterMassBalance : BOOL
VAR_INPUT
    rFeedM3h : REAL; // 进泥体积流量 [m3/h] / feed sludge flow
    rFeedTsPct : REAL; // 进泥含固率 [%] / feed total solids
    rCakeTsPct : REAL; // 泥饼含固率 [%] / cake total solids
    rFiltrateTsPct : REAL; // 滤液含固率 [%]，固体损失实测 / filtrate solids, measured loss
END_VAR
VAR_OUTPUT
    rCakeM3h : REAL; // 泥饼体积流量 [m3/h] / cake flow
    rFiltrateM3h : REAL; // 滤液体积流量 [m3/h] / filtrate flow
    rRecoveryPct : REAL; // 固体回收率 [%] / solids recovery
    bValid : BOOL; // 结果有效位 [-] / result valid flag
    iErrCode : INT; // 事件码 0=正常 1=泥饼含固率非法或不高於进泥 2=滤液量为负已归零 3=进泥流量非法 4=结果非有限 / event code
END_VAR
VAR CONSTANT
    rRecoveryCap : REAL := 100.0; // 回收率饱和上限 [%] / recovery saturation cap
END_VAR
VAR
    rCakeRaw : REAL; // 未校验泥饼量 [m3/h] / unchecked cake flow
    rFilRaw : REAL; // 未校验滤液量 [m3/h] / unchecked filtrate flow
    rFeedSolid : REAL; // 进泥固体负荷 [%·m3/h] / feed solids product
    rLossSolid : REAL; // 滤液固体损失 [%·m3/h] / filtrate solids loss
END_VAR

    // —— 段 0：全路径预清 —— //
    rCakeRaw := 0.0;
    rFilRaw := 0.0;
    rFeedSolid := 0.0;
    rCakeM3h := 0.0;
    rFiltrateM3h := 0.0;
    rRecoveryPct := 0.0;
    bValid := FALSE;
    iErrCode := 0;
    FC_DL_DewaterMassBalance := FALSE;
    // —— 段 1：分母闸与物理域闸（泥饼含固率必须高于进泥） —— //
    IF (rCakeTsPct <= 0.0) OR (rCakeTsPct <= rFeedTsPct) THEN
        iErrCode := 1; // 泥饼含固率非法或未脱水，平衡失效 / cake solids invalid or no dewatering achieved
        RETURN;
    END_IF;
    IF rFeedM3h <= 0.0 THEN
        iErrCode := 3; // 进泥流量非法 / invalid feed flow
        RETURN;
    END_IF;
    // —— 段 2：量纲链 (%·m3/h)/(%) = m3/h —— //
    rCakeRaw := rFeedM3h * rFeedTsPct / rCakeTsPct; // 泥饼量 [m3/h] / cake flow
    IF ABS(rCakeRaw) > 1.0E15 THEN
        iErrCode := 4; // 结果非有限，强制归零 / non-finite result, forced to zero
        RETURN;
    END_IF;
    rCakeM3h := rCakeRaw;
    // —— 段 3：滤液量 = 进泥量 - 泥饼量，负值归零并置码 —— //
    rFilRaw := rFeedM3h - rCakeM3h; // 滤液量 [m3/h] / filtrate flow
    IF rFilRaw < 0.0 THEN
        rFiltrateM3h := 0.0;
        iErrCode := 2; // 负滤液量（含固率组合不自洽）已归零 / negative filtrate clamped to zero
    ELSE
        rFiltrateM3h := rFilRaw;
    END_IF;
    // —— 段 4：回收率（分母闸：进泥固体负荷） —— //
    rFeedSolid := rFeedTsPct * rFeedM3h; // 进泥固体负荷 [%·m3/h] / feed solids
    IF ABS(rFeedSolid) <= 1.0E-9 THEN
        rRecoveryPct := 0.0; // 无固体，回收率无定义置零 / no solids, recovery undefined
    ELSE
        // 原式分子为平衡产物，恒等于 100%，改为按滤液损失实测
        IF rFiltrateTsPct < 0.0 THEN
            rFiltrateTsPct := 0.0; // 负含固率防御 / negative solids guard
        END_IF
        rLossSolid := rFiltrateTsPct * rFiltrateM3h; // 滤液带走固体 [%·m3/h] / lost solids
        rRecoveryPct := (rFeedSolid - rLossSolid) / rFeedSolid * 100.0; // 回收率 [%] / recovery by loss
        IF rRecoveryPct > rRecoveryCap THEN
            rRecoveryPct := rRecoveryCap; // 饱和 100% / saturate at 100 percent
        END_IF
    END_IF;
    bValid := TRUE;
    FC_DL_DewaterMassBalance := TRUE;
END_FUNCTION

(* ---- FC_DL_DiacetylRestWindowCalc.st ---- *)
// FC_DL_DiacetylRestWindowCalc v1.0.0
// 开源溯源：clean-room 自研（族 DL_Process，ST 生态实测 0 命中，无外部代码引入）
(*
  功能: 双乙酰还原时长：速率 = 参考速率·2^((T − Tref)/10)（Q10 = 2 工程近似，每升 10 °C 翻倍），
        时长 = LN(当前/目标)/速率 [h]；当前不高于目标时直接返回 0（已达标，不判错）。
  邻件/码位: 与 FC_DL_FermentAttenuationCalc 同属发酵后段件（主发酵终点 vs 还原终点）；
             16#0002_9236 = 非有限、浓度非正、参考速率非正或速率近零拒收。
*)
FUNCTION FC_DL_DiacetylRestWindowCalc : REAL
VAR_INPUT
    fTemp           : REAL := 14.0; // 还原温度 [°C] / Rest temperature [degC]
    fDiacetylNow    : REAL := 0.30; // 当前双乙酰 [mg/L]，域 > 0 / Current diacetyl [mg/L]
    fDiacetylTarget : REAL := 0.10; // 目标双乙酰 [mg/L]，域 > 0 / Target diacetyl [mg/L]
    fRateRef        : REAL := 0.05; // 参考温度衰减速率 [1/h]，域 > 0 / Decay rate at reference
    fTempRef        : REAL := 20.0; // 参考温度 [°C] / Reference temperature [degC]
END_VAR
VAR_OUTPUT
    fHoursNeeded : REAL;            // 预计还原时长 [h] / Estimated rest duration [h]
    bValid       : BOOL;            // 结果有效回执 [-] / Result validity receipt
    uErrorId     : UDINT;           // 事件码，0 = 无事件 / Event code
END_VAR
VAR
    fRate : REAL := 0.0;            // 实际衰减速率 [1/h] / Effective decay rate [1/h]
END_VAR
// 段 0：全路径出口安全缺省 / Safe defaults on all outlets
fHoursNeeded := 0.0;                // 时长缺省零 / Duration default zero
bValid := FALSE;                    // 有效回执预清 / Validity preset clear
uErrorId := 16#0000;                // 事件码预清 / Event code preset clear
FC_DL_DiacetylRestWindowCalc := 0.0;    // 返回值缺省零（镜像时长）/ Return default zero
// 段 1：非有限闸（五入参全枚举）/ Non-finite gate over all inputs
IF (fTemp <> fTemp) OR (fDiacetylNow <> fDiacetylNow) OR (fDiacetylTarget <> fDiacetylTarget)
   OR (fRateRef <> fRateRef) OR (fTempRef <> fTempRef)
   OR (ABS(fTemp) >= 3.0E38) OR (ABS(fDiacetylNow) >= 3.0E38) OR (ABS(fDiacetylTarget) >= 3.0E38)
   OR (ABS(fRateRef) >= 3.0E38) OR (ABS(fTempRef) >= 3.0E38) THEN
    uErrorId := 16#0002_9236;   // 入参非有限拒收 / Non-finite input reject
    RETURN;
END_IF
// 段 2：域闸（浓度与参考速率非正拒收 + 已达标快通道，R4）/ Domain gate
IF (fDiacetylNow <= 0.0) OR (fDiacetylTarget <= 0.0) THEN
    uErrorId := 16#0002_9236;   // 浓度非正，LN 无意义 / Non-positive concentration
    RETURN;
END_IF
IF fRateRef <= 1.0E-6 THEN
    uErrorId := 16#0002_9236;   // 参考速率非正 / Non-positive reference rate
    RETURN;
END_IF
IF fDiacetylNow <= fDiacetylTarget THEN
    bValid := TRUE;             // 已达标：时长零，仍为有效解 / Already compliant, valid
    RETURN;                     // 时长已由段 0 置零 / Duration stays zero from stage 0
END_IF
// 段 3：主计算（Q10 温度修正 → LN 比值 → 时长）/ Main computation
fRate := fRateRef * EXP((fTemp - fTempRef) / 10.0 * 0.693147180559945);     // ref·2^expo [1/h] / Effective rate
IF fRate <= 1.0E-9 THEN
    uErrorId := 16#0002_9236;   // 速率近零，时长发散 / Rate too small, duration diverges
    RETURN;
END_IF
fHoursNeeded := LN(fDiacetylNow / fDiacetylTarget) / fRate;     // 时长 [h] / Rest duration
// 段 4：出口闸（非有限复核 + 非负复核）/ Outlet gate
IF (fHoursNeeded <> fHoursNeeded) OR (ABS(fHoursNeeded) >= 3.0E38) OR (fHoursNeeded < 0.0) THEN
    fHoursNeeded := 0.0;        // 复核失败回缺省 / Fallback on recheck failure
    uErrorId := 16#0002_9236;   // 出口复核拒收 / Output recheck reject
    RETURN;
END_IF
bValid := TRUE;                 // 有效回执 / Validity receipt
FC_DL_DiacetylRestWindowCalc := fHoursNeeded;   // 返回值镜像时长 / Return mirrors duration
END_FUNCTION

(* ---- FC_DL_DieCastIntensifyPressureCalc.st ---- *)
(*
  Component : FC_DL_DieCastIntensifyPressureCalc
  Category  : DL_Process
  Type      : FC
  Complexity: C2
  VERSION   : v1.0.0
  功能      : 增压比压与锁模力校验：按铸件投影面积与增压比压算所需锁模力，并与设备额定锁模力比较输出余量比。
  开源溯源  : 道莅原创 clean-room 自研（无外部代码引用）｜License: MIT
  边界条件  : ① 投影面积、增压比压、安全系数须 > 1e-9，否则返回哨兵 -1；
              ② 所需锁模力 = 投影面积(cm²) × 比压(MPa) / 10 × 安全系数，量纲为 kN；
              ③ 余量比 = 额定/所需，额定为 0 时不计算而回哨兵。
*)
FUNCTION FC_DL_DieCastIntensifyPressureCalc : REAL
VAR_INPUT
    fProjAreaCm2    : REAL;   (* 铸件投影面积（含浇排系统） [cm²] Projected area *)
    fCastPressMPa   : REAL;   (* 压射比压 [MPa] Casting specific pressure *)
    fIntensifyRatio : REAL;   (* 增压比（增压后/压射） [-] Intensification ratio *)
    fRatedClampKN   : REAL;   (* 设备额定锁模力 [kN] Rated clamping force *)
    fSafetyFactor   : REAL;   (* 锁模安全系数 [-] Clamping safety factor *)
END_VAR
VAR_OUTPUT
    fIntPressMPa  : REAL;  (* 增压后比压 [MPa] Intensified specific pressure *)
    fClampNeedKN  : REAL;  (* 所需锁模力 [kN] Required clamping force *)
    fMarginRatio  : REAL;  (* 锁模力余量比（额定/所需） [-] Clamping margin ratio *)
    xClampOk      : BOOL;  (* 锁模力充足标志 [-] Clamping sufficient flag *)
    xValid        : BOOL;  (* 计算有效性标志 [-] Calculation valid flag *)
END_VAR
VAR CONSTANT
    DL_EPS      : REAL := 1.0E-9;   (* 除零判定容差 [无量纲] Divide-by-zero tolerance *)
    DL_KPA_UNIT : REAL := 10.0;     (* cm²×MPa 换算 kN 的除数 [cm²·MPa/kN] Unit divisor *)
    DL_ZERO     : REAL := 0.0;      (* 零常量 [无量纲] Zero constant *)
END_VAR
(* 出口预置：五出口统一预置 *)
fIntPressMPa := 0.0; fClampNeedKN := 0.0; fMarginRatio := 0.0; xClampOk := FALSE; xValid := FALSE;
(* 非有限拦截：自反判 NaN，自身差值判 Inf *)
IF (fProjAreaCm2 <> fProjAreaCm2) OR ((fProjAreaCm2 - fProjAreaCm2) <> 0.0)
   OR (fCastPressMPa <> fCastPressMPa) OR ((fCastPressMPa - fCastPressMPa) <> 0.0)
   OR (fIntensifyRatio <> fIntensifyRatio) OR ((fIntensifyRatio - fIntensifyRatio) <> 0.0)
   OR (fRatedClampKN <> fRatedClampKN) OR ((fRatedClampKN - fRatedClampKN) <> 0.0)
   OR (fSafetyFactor <> fSafetyFactor) OR ((fSafetyFactor - fSafetyFactor) <> 0.0) THEN
    FC_DL_DieCastIntensifyPressureCalc := -1.0;  (* 哨兵 -1：输入非有限 / Sentinel -1 non-finite *)
    RETURN;
END_IF
(* 组态域闸：面积、比压、增压比、安全系数、额定锁模力逐个覆盖 *)
IF (fProjAreaCm2 <= DL_EPS) OR (fCastPressMPa <= DL_ZERO) OR (fIntensifyRatio <= DL_EPS)
   OR (fSafetyFactor <= DL_EPS) OR (fRatedClampKN <= DL_ZERO) THEN
    FC_DL_DieCastIntensifyPressureCalc := -1.0;  (* 哨兵 -1：组态非法 / Sentinel -1 bad config *)
    RETURN;
END_IF
(* 增压后比压：p2 = p × 增压比 [MPa] *)
fIntPressMPa := fCastPressMPa * fIntensifyRatio;
(* 所需锁模力：A(cm²)=100 mm²，p(MPa)=N/mm²，F=100·A·p N = A·p/10 kN *)
fClampNeedKN := fProjAreaCm2 * fIntPressMPa / DL_KPA_UNIT * fSafetyFactor;
(* 余量比：额定 / 所需，所需已过域闸（面积与比压均正） *)
fMarginRatio := fRatedClampKN / fClampNeedKN;
xClampOk := fMarginRatio >= 1.0;                (* 余量比 >= 1 判充足 / Sufficient margin *)
xValid := TRUE;                                 (* 链路有效 / Chain valid *)
FC_DL_DieCastIntensifyPressureCalc := fClampNeedKN;  (* 返回所需锁模力 [kN] / Return clamp force *)
END_FUNCTION

(* ---- FC_DL_DieCastShotVelocityCalc.st ---- *)
(*
  Component : FC_DL_DieCastShotVelocityCalc
  Category  : DL_Process
  Type      : FC
  Complexity: C2
  VERSION   : v1.0.0
  功能      : 压射速度核算：按充填体积/充填时间/冲头面积算空压射速度，做 PQ² 交点速度校核并给出超限降速建议。
  开源溯源  : 道莅原创 clean-room 自研（无外部代码引用）｜License: MIT
  边界条件  : ① 充填时间、冲头直径、充填体积须 > 1e-9，否则返回哨兵 -1（充填时间为除子）；
              ② 速度超工艺上限置 xOverLimit；速度超 PQ² 交点速度置 xPq2Ok = FALSE 并给降速建议；
              ③ 降速建议 = min(0.9 × PQ² 交点速度, 工艺上限)，不越上限。
*)
FUNCTION FC_DL_DieCastShotVelocityCalc : REAL
VAR_INPUT
    fFillVolCm3   : REAL;   (* 型腔充填体积 [cm³] Cavity fill volume *)
    fFillTimeMs   : REAL;   (* 充填时间 [ms] Fill time *)
    fPlungerDiaMm : REAL;   (* 压射冲头直径 [mm] Shot plunger diameter *)
    fMaxVelMs     : REAL;   (* 工艺允许最大速度 [m/s] Process max velocity *)
    fPq2VelMs     : REAL;   (* PQ² 交点速度 [m/s] PQ2 intersection velocity *)
END_VAR
VAR_OUTPUT
    fShotVelMs   : REAL;  (* 空压射速度 [m/s] Dry shot velocity *)
    fPq2Ratio    : REAL;  (* 速度 / PQ² 交点速度比 [-] Velocity to PQ2 ratio *)
    fSuggestVelMs: REAL;  (* 超限降速建议值 [m/s] Suggested reduced velocity *)
    xOverLimit   : BOOL;  (* 超工艺上限标志 [-] Over process limit flag *)
    xPq2Ok       : BOOL;  (* PQ² 校核通过标志 [-] PQ2 check passed flag *)
    xValid       : BOOL;  (* 计算有效性标志 [-] Calculation valid flag *)
END_VAR
VAR CONSTANT
    DL_EPS      : REAL := 1.0E-9;   (* 除零判定容差 [无量纲] Divide-by-zero tolerance *)
    DL_PI       : REAL := 3.14159265358979;  (* 圆周率 [-] Pi *)
    DL_MS_PER_S : REAL := 1000.0;   (* 毫秒转秒换算系数 [ms/s] Milliseconds per second *)
    DL_SAFE_K   : REAL := 0.9;      (* 降速安全系数 [-] Velocity reduction factor *)
    DL_ZERO     : REAL := 0.0;      (* 零常量 [无量纲] Zero constant *)
END_VAR
VAR
    fAreaMm2 : REAL;   (* 冲头截面积 [mm²] Plunger cross-section *)
    fTimeS   : REAL;   (* 充填时间秒值 [s] Fill time in seconds *)
    fVelCm   : REAL;   (* 中间速度量 [cm³/(mm²·s)] Intermediate velocity *)
    fCand    : REAL;   (* 降速候选值 [m/s] Candidate reduced velocity *)
END_VAR
(* 出口预置：六出口统一预置 *)
fShotVelMs := 0.0; fPq2Ratio := 0.0; fSuggestVelMs := 0.0;
xOverLimit := FALSE; xPq2Ok := FALSE; xValid := FALSE;
(* 非有限拦截：自反判 NaN，自身差值判 Inf *)
IF (fFillVolCm3 <> fFillVolCm3) OR ((fFillVolCm3 - fFillVolCm3) <> 0.0)
   OR (fFillTimeMs <> fFillTimeMs) OR ((fFillTimeMs - fFillTimeMs) <> 0.0)
   OR (fPlungerDiaMm <> fPlungerDiaMm) OR ((fPlungerDiaMm - fPlungerDiaMm) <> 0.0)
   OR (fMaxVelMs <> fMaxVelMs) OR ((fMaxVelMs - fMaxVelMs) <> 0.0)
   OR (fPq2VelMs <> fPq2VelMs) OR ((fPq2VelMs - fPq2VelMs) <> 0.0) THEN
    FC_DL_DieCastShotVelocityCalc := -1.0;  (* 哨兵 -1：输入非有限 / Sentinel -1 non-finite *)
    RETURN;
END_IF
(* 组态域闸：体积/时间/直径为除子，两个速度限须为正 *)
IF (fFillVolCm3 <= DL_EPS) OR (fFillTimeMs <= DL_EPS) OR (fPlungerDiaMm <= DL_EPS)
   OR (fMaxVelMs <= DL_ZERO) OR (fPq2VelMs <= DL_ZERO) THEN
    FC_DL_DieCastShotVelocityCalc := -1.0;  (* 哨兵 -1：组态非法 / Sentinel -1 bad config *)
    RETURN;
END_IF
fAreaMm2 := DL_PI / 4.0 * fPlungerDiaMm * fPlungerDiaMm;   (* 冲头面积 [mm²] *)
fTimeS := fFillTimeMs / DL_MS_PER_S;                       (* 充填时间 [s] *)
(* 速度换算：cm³/(mm²·s) = 1000 mm³/(mm²·s) = 1000 mm/s = 1 m/s，故量纲直接得 m/s *)
fVelCm := fFillVolCm3 / (fAreaMm2 * fTimeS);
fShotVelMs := fVelCm;
(* PQ² 校核：速度比与通过标志 *)
fPq2Ratio := fShotVelMs / fPq2VelMs;
xPq2Ok := fShotVelMs <= fPq2VelMs;
xOverLimit := fShotVelMs > fMaxVelMs;
(* 降速建议：取 0.9 倍 PQ² 交点速度与工艺上限的较小者 *)
IF xOverLimit OR (NOT xPq2Ok) THEN
    fCand := fPq2VelMs * DL_SAFE_K;
    IF fCand < fMaxVelMs THEN
        fSuggestVelMs := fCand;                 (* 受 PQ² 交点约束 [m/s] / Limited by PQ2 *)
    ELSE
        fSuggestVelMs := fMaxVelMs;             (* 受工艺上限约束 [m/s] / Limited by process cap *)
    END_IF
ELSE
    fSuggestVelMs := fShotVelMs;                (* 未超限：建议保持当前速度 *)
END_IF
xValid := TRUE;                                 (* 链路有效 / Chain valid *)
FC_DL_DieCastShotVelocityCalc := fShotVelMs;    (* 返回空压射速度 [m/s] / Return shot velocity *)
END_FUNCTION

(* ---- FC_DL_DieThermalBalanceCalc.st ---- *)
(*
  Component : FC_DL_DieThermalBalanceCalc
  Category  : DL_Process
  Type      : FC
  Complexity: C2
  VERSION   : v1.0.0
  功能      : 压铸模热平衡核算：按循环周期与金属放热算平均热流，再由冷却水流量算水温升与模温估计，给出模温机负荷。
  开源溯源  : 道莅原创 clean-room 自研（无外部代码引用）｜License: MIT
  边界条件  : ① 循环周期、金属质量、比热、冷却水流量均须 > 1e-9，否则返回哨兵 -1；
              ② 放热按金属从浇注温度降到顶出温度的显热估算，不含凝固潜热；
              ③ 浇注温度低于顶出温度时放热量归零；模温机余量上限钳位 100 %（折算系数上限 2.0）。
*)
FUNCTION FC_DL_DieThermalBalanceCalc : REAL
VAR_INPUT
    fCycleS       : REAL;   (* 压铸循环周期 [s] Die casting cycle time *)
    fMetalMassKg  : REAL;   (* 单模金属质量 [kg] Metal mass per shot *)
    fMetalCpKJkgK : REAL;   (* 金属比热容 [kJ/(kg·K)] Metal specific heat *)
    fPourC        : REAL;   (* 浇注温度 [°C] Pouring temperature *)
    fEjectC       : REAL;   (* 顶出温度 [°C] Ejection temperature *)
    fWaterFlowLmin: REAL;   (* 冷却水流量 [L/min] Cooling water flow *)
    fWaterInC     : REAL;   (* 冷却水进水温度 [°C] Cooling water inlet temperature *)
    fMarginPct    : REAL;   (* 模温机负荷余量 [%] Thermolator load margin *)
END_VAR
VAR_OUTPUT
    fHeatRateKW  : REAL;  (* 模具平均热流 [kW] Average heat flux into die *)
    fCoolLoadKW  : REAL;  (* 模温机所需冷却负荷 [kW] Required cooling load *)
    fWaterDeltaTK: REAL;  (* 冷却水温升 [K] Cooling water temperature rise *)
    fMoldEstC    : REAL;  (* 模温估计 [°C] Estimated die temperature *)
    xValid       : BOOL;  (* 计算有效性标志 [-] Calculation valid flag *)
END_VAR
VAR CONSTANT
    DL_EPS      : REAL := 1.0E-9;   (* 除零判定容差 [无量纲] Divide-by-zero tolerance *)
    DL_S_PER_MIN: REAL := 60.0;     (* 分钟转秒换算系数 [s/min] Seconds per minute *)
    DL_WATER_CP : REAL := 4.187;    (* 水比热容 [kJ/(kg·K)] Water specific heat *)
    DL_PCT_BASE : REAL := 100.0;    (* 百分比基准 [%] Percent base *)
    DL_ZERO     : REAL := 0.0;      (* 零常量 [无量纲] Zero constant *)
END_VAR
VAR
    fHeatKJ    : REAL;   (* 单模放热量 [kJ] Heat per shot *)
    fFlowKgS   : REAL;   (* 冷却水质量流量 [kg/s] Cooling water mass flow *)
    fMarginK   : REAL;   (* 余量折算系数 [-] Margin factor *)
END_VAR
(* 出口预置：五出口统一预置 *)
fHeatRateKW := 0.0; fCoolLoadKW := 0.0; fWaterDeltaTK := 0.0; fMoldEstC := 0.0; xValid := FALSE;
(* 非有限拦截：自反判 NaN，自身差值判 Inf *)
IF (fCycleS <> fCycleS) OR ((fCycleS - fCycleS) <> 0.0)
   OR (fMetalMassKg <> fMetalMassKg) OR ((fMetalMassKg - fMetalMassKg) <> 0.0)
   OR (fMetalCpKJkgK <> fMetalCpKJkgK) OR ((fMetalCpKJkgK - fMetalCpKJkgK) <> 0.0)
   OR (fPourC <> fPourC) OR ((fPourC - fPourC) <> 0.0)
   OR (fEjectC <> fEjectC) OR ((fEjectC - fEjectC) <> 0.0)
   OR (fWaterFlowLmin <> fWaterFlowLmin) OR ((fWaterFlowLmin - fWaterFlowLmin) <> 0.0)
   OR (fWaterInC <> fWaterInC) OR ((fWaterInC - fWaterInC) <> 0.0)
   OR (fMarginPct <> fMarginPct) OR ((fMarginPct - fMarginPct) <> 0.0) THEN
    FC_DL_DieThermalBalanceCalc := -1.0;  (* 哨兵 -1：输入非有限 / Sentinel -1 non-finite *)
    RETURN;
END_IF
(* 组态域闸：周期、质量、比热为比例基；流量为水温升的除子 *)
IF (fCycleS <= DL_EPS) OR (fMetalMassKg <= DL_EPS) OR (fMetalCpKJkgK <= DL_EPS)
   OR (fWaterFlowLmin <= DL_EPS) OR (fMarginPct < DL_ZERO) THEN
    FC_DL_DieThermalBalanceCalc := -1.0;  (* 哨兵 -1：组态非法 / Sentinel -1 bad config *)
    RETURN;
END_IF
(* 单模显热：Q = m·cp·ΔT [kJ]，ΔT 为浇注与顶出温差 *)
fHeatKJ := fMetalMassKg * fMetalCpKJkgK * (fPourC - fEjectC);
IF fHeatKJ < DL_ZERO THEN
    fHeatKJ := DL_ZERO;                       (* 负温差归零 [kJ] / Negative heat clamp *)
END_IF
(* 平均热流：Q / 周期 [kJ/s = kW] *)
fHeatRateKW := fHeatKJ / fCycleS;
(* 模温机负荷：平均热流 × (1 + 余量)，余量钳位 0~100 % *)
fMarginK := 1.0 + fMarginPct / DL_PCT_BASE;
IF fMarginK > 2.0 THEN
    fMarginK := 2.0;                          (* 余量上限钳位 [-] / Margin upper clamp *)
END_IF
fCoolLoadKW := fHeatRateKW * fMarginK;
(* 水温升：Q = m·cp·ΔT，水质量流量 L/min ÷ 60 = kg/s，分母已过域闸 *)
fFlowKgS := fWaterFlowLmin / DL_S_PER_MIN;
fWaterDeltaTK := fHeatRateKW / (fFlowKgS * DL_WATER_CP);
(* 模温估计：进水温度叠加水温升（模具侧平均近似） *)
fMoldEstC := fWaterInC + fWaterDeltaTK;
xValid := TRUE;                               (* 链路有效 / Chain valid *)
FC_DL_DieThermalBalanceCalc := fCoolLoadKW;   (* 返回冷却负荷 [kW] / Return cooling load *)
END_FUNCTION

(* ---- FC_DL_DigesterRetentionTime.st ---- *)
(*
  道莅工业代码库 / Daoli Industrial ST Library
  组件: FC_DL_DigesterRetentionTime
  分类: DL_Process
  开源溯源: 无（clean-room 工程公式自研；参考公开工艺计算公式，未复制任何受版权保护代码）
  许可证: 本项目自有 (MIT)
  功能: 消化罐水力停留时间 HRT、固体停留时间 SRT 与容积负荷估算
  口径声明: 容积负荷按进料 VS 浓度假定 25 kg/m3 折算（现场标定前作为默认口径），
            SRT 分母取「废弃污泥流量 + 进料量的 2%（随出流带出固体）」
*)
FUNCTION FC_DL_DigesterRetentionTime : BOOL
VAR_INPUT
    rReactorM3 : REAL; // 反应器有效容积 [m3] / reactor working volume
    rFeedM3Day : REAL; // 进料流量 [m3/d] / feed flow
    rRecycleM3Day : REAL; // 废弃污泥（排泥）流量 [m3/d] / waste sludge flow
END_VAR
VAR_OUTPUT
    rHrtDay : REAL; // 水力停留时间 [d] / hydraulic retention time
    rSrtDay : REAL; // 固体停留时间 [d] / solids retention time
    rLoadingKgM3d : REAL; // 容积有机负荷 [kgVS/(m3·d)] / volumetric organic loading
    bValid : BOOL; // 结果有效位 [-] / result valid flag
    iErrCode : INT; // 事件码 0=正常 1=进料流量非法 2=SRT 小于 HRT 已按 HRT 饱和 3=结果非有限 / event code
END_VAR
VAR CONSTANT
    rVsConcAssumed : REAL := 25.0; // 进料 VS 浓度假定值 [kgVS/m3] / assumed feed VS concentration
    rCarryFrac : REAL := 0.02; // 出流带出固体占进料比 [-] / solids carry-out fraction of feed
END_VAR
VAR
    rQTotalM3d : REAL; // 总吞吐流量 [m3/d] / total through flow
    rQOutM3d : REAL; // 固体出流当量流量 [m3/d] / solids outflow equivalent
    rHrtRaw : REAL; // 未校验 HRT [d] / unchecked HRT
    rSrtRaw : REAL; // 未校验 SRT [d] / unchecked SRT
    rLoadingRaw : REAL; // 未校验负荷 [kgVS/(m3·d)] / unchecked loading
END_VAR

    // —— 段 0：全路径预清 —— //
    rQTotalM3d := 0.0;
    rQOutM3d := 0.0;
    rHrtRaw := 0.0;
    rSrtRaw := 0.0;
    rLoadingRaw := 0.0;
    rHrtDay := 0.0;
    rSrtDay := 0.0;
    rLoadingKgM3d := 0.0;
    bValid := FALSE;
    iErrCode := 0;
    FC_DL_DigesterRetentionTime := FALSE;
    // —— 段 1：分母闸（总吞吐流量 = 进料 + 回流/排泥） —— //
    rQTotalM3d := rFeedM3Day + rRecycleM3Day; // 总吞吐 [m3/d] / total through flow
    IF (rQTotalM3d <= 0.0) OR (rFeedM3Day <= 0.0) THEN
        iErrCode := 1; // 流量非法，停留时间无定义 / invalid flow, retention time undefined
        RETURN;
    END_IF;
    IF rReactorM3 <= 0.0 THEN
        iErrCode := 1; // 容积非法 / invalid volume
        RETURN;
    END_IF;
    // —— 段 2：量纲链 (m3)/(m3/d) = d —— //
    rHrtRaw := rReactorM3 / rQTotalM3d; // HRT [d] / hydraulic retention time
    IF ABS(rHrtRaw) > 1.0E15 THEN
        iErrCode := 3; // 结果非有限，强制归零 / non-finite result, forced to zero
        RETURN;
    END_IF;
    rHrtDay := rHrtRaw;
    // —— 段 3：SRT 分母 = 排泥量 + 进料×2%（分母闸：不得为零） —— //
    rQOutM3d := rRecycleM3Day + rFeedM3Day * rCarryFrac; // 固体出流当量 [m3/d] / solids outflow equivalent
    IF rQOutM3d <= 1.0E-9 THEN
        rSrtDay := rHrtDay; // 无排泥即无固体流出，SRT 退化按 HRT 计 / no wasting, SRT falls back to HRT
        iErrCode := 2; // 信息级：SRT 按 HRT 饱和 / info level: SRT saturated at HRT
    ELSE
        rSrtRaw := rReactorM3 / rQOutM3d; // SRT [d] / solids retention time
        IF ABS(rSrtRaw) > 1.0E15 THEN
            rSrtRaw := rHrtDay; // 非有限兜底 / non-finite fallback
            iErrCode := 3;
        END_IF;
        IF rSrtRaw < rHrtDay THEN
            rSrtDay := rHrtDay; // SRT 不可能小于 HRT，饱和到 HRT / SRT cannot be below HRT
            iErrCode := 2; // 信息级：SRT 参数不自洽 / info level: SRT parameters inconsistent
        ELSE
            rSrtDay := rSrtRaw;
        END_IF
    END_IF;
    // —— 段 4：容积负荷（量纲 (m3/d)×(kg/m3)/(m3) = kg/(m3·d)） —— //
    rLoadingRaw := rFeedM3Day * rVsConcAssumed / rReactorM3; // 容积负荷 [kgVS/(m3·d)] / volumetric loading
    IF ABS(rLoadingRaw) > 1.0E15 THEN
        rLoadingKgM3d := 0.0;
        iErrCode := 3; // 结果非有限，强制归零 / non-finite result, forced to zero
        RETURN;
    END_IF;
    rLoadingKgM3d := rLoadingRaw;
    bValid := TRUE;
    FC_DL_DigesterRetentionTime := TRUE;
END_FUNCTION

(* ---- FC_DL_DoDeficitCalc.st ---- *)
(*
  ============================================================
  组件名 : FC_DL_DoDeficitCalc
  分类   : DL_Process
  功能   : 溶解氧偏差与饱和度计算，按实测值与设定值求欠氧量并双向分档
  开源溯源 : internal-design（本轮无外部代码逐行引用）
             参考语义 : 无外部参考
  复杂度 : C1
  版本   : 1.0.0
  ============================================================
*)

FUNCTION FC_DL_DoDeficitCalc : REAL
VAR_INPUT
    rDoAct_mgL : REAL; // 实测溶解氧 [mg/L] measured dissolved oxygen [mg per litre]
    rDoSp_mgL  : REAL; // 溶解氧设定值 [mg/L] dissolved oxygen set point [mg per litre]
    rDoLow     : REAL; // 偏低判定阈值 [mg/L] low verdict threshold [mg per litre]
    rDoHigh    : REAL; // 偏高判定阈值 [mg/L] high verdict threshold [mg per litre]
END_VAR
VAR_OUTPUT
    rDeficit       : REAL; // 溶解氧欠量，设定减实测 [mg/L] oxygen deficit, set point minus actual [mg per litre]
    rSaturationPct : REAL; // 实测相对设定的百分比 [%] actual relative to the set point [%]
    nStatus        : INT; // 分档 0正常 1偏低 2偏高 [档] status 0 normal, 1 low, 2 high [band]
    bValid         : BOOL; // 结果有效标志 result validity flag
END_VAR
VAR CONSTANT
    DL_HUNDRED : REAL := 100.0; // 百分制换算系数 percentage scale factor
    DL_EPS_R   : REAL := 1.0E-6; // 实数零判定阈值 real zero threshold
END_VAR
VAR
    _bFin : BOOL := FALSE; // 四输入有限性判定 finiteness verdict of the four inputs
    _rDef : REAL := 0.0; // 欠量中间量 [mg/L] intermediate deficit [mg per litre]
    _rSat : REAL := 0.0; // 百分比中间量 [%] intermediate percentage [%]
    _rLow : REAL := 0.0; // 钳位后的偏低阈值 [mg/L] clamped low threshold [mg per litre]
    _rHigh: REAL := 0.0; // 钳位后的偏高阈值 [mg/L] clamped high threshold [mg per litre]
END_VAR

// 段 1｜出口预置 preset the exit
FC_DL_DoDeficitCalc := 0.0; // 缺省返回零 default zero return
rDeficit := 0.0; // 欠量预置零 deficit preset to zero
rSaturationPct := 0.0; // 百分比预置零 percentage preset to zero
nStatus := 0; // 分档预置正常 status preset normal
bValid := FALSE; // 计算完成前不认结果 unusable before the calculation
// 段 2｜非有限闸 finiteness gate
_bFin := (rDoAct_mgL = rDoAct_mgL) AND (rDoSp_mgL = rDoSp_mgL) AND (rDoLow = rDoLow) AND (rDoHigh = rDoHigh); // 四输入自反判定 self comparison of the four inputs
IF NOT _bFin THEN
    RETURN; // 非有限即无效 non finite means invalid
END_IF
// 段 3｜设定值分母闸 set point divisor gate
IF rDoSp_mgL <= DL_EPS_R THEN
    RETURN; // 设定值非正无法折算百分比 a non positive set point cannot carry a percentage
END_IF
// 段 4｜欠量与百分比 deficit and the percentage
_rDef := rDoSp_mgL - rDoAct_mgL; // 设定减实测 set point minus actual
_rSat := rDoAct_mgL / rDoSp_mgL * DL_HUNDRED; // 实测占设定百分比 actual over the set point
rDeficit := _rDef; // 欠量落定 land the deficit
rSaturationPct := _rSat; // 百分比落定 land the percentage
// 段 5｜双向分档判定 directional status verdict
_rLow := rDoLow; // 取偏低阈值 take the low threshold
_rHigh := rDoHigh; // 取偏高阈值 take the high threshold
IF _rLow > _rHigh THEN
    _rLow := rDoHigh; // 阈值倒置时偏低阈值取原偏高 an inverted pair swaps the low threshold
    _rHigh := rDoLow; // 阈值倒置时偏高阈值取原偏低 an inverted pair swaps the high threshold
END_IF
IF rDoAct_mgL < _rLow THEN
    nStatus := 1; // 实测偏低 the reading is too low
ELSIF rDoAct_mgL > _rHigh THEN
    nStatus := 2; // 实测偏高 the reading is too high
ELSE
    nStatus := 0; // 区间内正常 inside the normal band
END_IF
bValid := TRUE; // 结果可用 result usable
FC_DL_DoDeficitCalc := _rDef; // 函数返回欠量 return the deficit
END_FUNCTION

(* ---- FC_DL_DrainIntervalCalc.st ---- *)
(*
  ============================================================
  组件名 : FC_DL_DrainIntervalCalc
  分类   : DL_Process
  功能   : 自动排水间隔计算，由冷凝析水率与允许最大积水求排水周期并给出即时排水请求
  复杂度 : C1
  版本   : 1.0.0
  作者   : 道莅工业代码库工厂 / R81
  日期   : 2026-11-24
  开源溯源 : clean-room（no upstream）—— 依据公开工程公式自研，未复制任何上游实现
  红线自检 : R1 无GVL/R2 无物理地址/R3 纯IEC/R4 防除零/R5 双语注释
  接口说明 :
      排水间隔 = 允许最大积水 / 析水率 * 60，单位 min。
      间隔小于 10 min 表示积水速度已超出常规排放节奏，置 bDrainNow 请求连续排放。
      单次排水量仅用于校核排放能力是否覆盖间隔内的积水，不参与间隔公式。
  ============================================================
*)
FUNCTION FC_DL_DrainIntervalCalc : BOOL
VAR_INPUT
    bEnable      : BOOL; // 使能：TRUE 时计算 / Enable: TRUE to compute
    bErr         : BOOL; // 外部故障：TRUE 时立即退出并置结果无效 / External fault: TRUE aborts with invalid result
    rCondRate    : REAL; // 冷凝析水率 [L/h] / condensate generation rate [litre per hour]
    rDrainVol_L  : REAL; // 单次排水动作排放量 [L] / volume released by one drain action [litre]
    rMaxHold_L   : REAL; // 允许的最大积水量 [L] / maximum permitted accumulated water [litre]
END_VAR
VAR_OUTPUT
    rInterval_min : REAL; // 建议排水间隔 [min] / recommended drain interval [minute]
    rWaterPerInt_L : REAL; // 单个间隔内积水总量 [L] / accumulated water within one interval [litre]
    bDrainNow   : BOOL; // 即时排水请求：TRUE 表示间隔小于 10 min / immediate drain request, TRUE when the interval is below 10 minutes
    bCapOk      : BOOL; // 排放能力充足：TRUE 表示单次排放量不小于间隔内积水量 / capacity adequate, TRUE when one drain covers the water of one interval
    bValid      : BOOL; // 输出有效：TRUE 表示结果可用 / Output valid
END_VAR
VAR CONSTANT
    DL_R_MAX    : REAL := 3.0E38; // 实数上界，用于拦截 Inf [无量纲] / real upper bound used to reject infinity [dimensionless]
    DL_EPS      : REAL := 1.0E-12; // 除零判定阈值 [无量纲] / division guard threshold [dimensionless]
    DL_MIN_PER_H : REAL := 60.0;  // 每小时分钟数 [min/h] / minutes per hour [minute per hour]
    DL_NOW_MIN  : REAL := 10.0;   // 即时排水间隔门限 [min] / threshold of the immediate drain interval [minute]
    DL_TOL_L    : REAL := 1.0E-6; // 排放能力比较容差 [L] / tolerance of the drain capacity comparison [litre]
END_VAR
VAR
    _bFin : BOOL := FALSE; // 输入有限性判定结果 / input finiteness verdict
END_VAR

    // 段 1｜出口预置
    rInterval_min := 0.0;
    rWaterPerInt_L := 0.0;
    bDrainNow := FALSE;
    bCapOk := FALSE;
    bValid := FALSE;
    // 段 2｜使能闸与外部故障闸
    IF NOT bEnable THEN
        RETURN;
    END_IF;
    IF bErr THEN
        RETURN;
    END_IF;
    // 段 3｜非有限闸
    _bFin := (rCondRate = rCondRate) AND (ABS(rCondRate) <= DL_R_MAX) AND (rDrainVol_L = rDrainVol_L) AND (ABS(rDrainVol_L) <= DL_R_MAX) AND (rMaxHold_L = rMaxHold_L) AND (ABS(rMaxHold_L) <= DL_R_MAX);
    IF NOT _bFin THEN
        RETURN;
    END_IF;
    // 段 4｜域闸：析水率严格为正，积水量与单次排放量不得为负
    IF (ABS(rCondRate) <= DL_EPS) OR (rCondRate < 0.0) THEN
        RETURN;
    END_IF;
    IF (rMaxHold_L < 0.0) OR (rDrainVol_L < 0.0) THEN
        RETURN;
    END_IF;
    // 段 5｜排水间隔
    rInterval_min := rMaxHold_L / rCondRate * DL_MIN_PER_H;
    // 段 6｜间隔内积水量
    rWaterPerInt_L := rCondRate * rInterval_min / DL_MIN_PER_H;
    // 段 7｜排放能力校核：单次排放量须覆盖一个间隔的积水
    IF rDrainVol_L >= (rWaterPerInt_L - DL_TOL_L) THEN
        bCapOk := TRUE;
    ELSE
        bCapOk := FALSE;
    END_IF;
    // 段 8｜即时排水请求
    IF rInterval_min < DL_NOW_MIN THEN
        bDrainNow := TRUE;
    ELSE
        bDrainNow := FALSE;
    END_IF;
    bValid := TRUE;
    FC_DL_DrainIntervalCalc := bValid;
END_FUNCTION

(* ---- FC_DL_DryerMoistureRemovalCalc.st ---- *)
(*
 * FC_DL_DryerMoistureRemovalCalc | C2 | DL_Process
 * 功能：烘丝机水分去除量与干物料流量（按进出口含水率，湿基）       单位：流量 [kg/h]、含水率 [%]
 * 工况边界：含水率须在 0~100 % 且出口 <100 %（入分母）；出口含水率应小于入口，否则去水量为负（回潮工况）时按 0 处理并置 xValid=TRUE（数值合法但非烘干）；仅干基不变量成立，不含热耗与风量
 * 代数值回代：G=5000 kg/h、w1=18 %、w2=12 % → Gd=5000×82/100=4100 kg/h、W=4100×6/88=279.5 kg/h（与 spec 回代行一致）
 * 开源溯源：clean-room 自研，未复制任何第三方代码（无外部来源）
 *)
FUNCTION FC_DL_DryerMoistureRemovalCalc : BOOL
VAR_INPUT
    rFeedKgH     : REAL := 5000.0;   // 入口湿基流量 | inlet wet basis mass flow [kg/h]
    rMoistInPct  : REAL := 18.0;     // 入口含水率（湿基）| inlet moisture, wet basis [%]
    rMoistOutPct : REAL := 12.0;     // 出口含水率（湿基）| outlet moisture, wet basis [%]
END_VAR
VAR_OUTPUT
    rWaterRemovedKgH : REAL;         // 去水量 | water removed [kg/h]
    rDryMatterKgH    : REAL;         // 绝干物料流量 | dry matter mass flow [kg/h]
    xReverseMoist    : BOOL;         // 出口含水率高于入口（回潮工况，信息级）| outlet moisture above the inlet, informational
    xValid           : BOOL;         // 输出有效 | outputs valid
END_VAR
VAR
    xFinG  : BOOL;                   // 入口流量有限性 | inlet flow is finite
    xFinW1 : BOOL;                   // 入口水分有限性 | inlet moisture is finite
    xFinW2 : BOOL;                   // 出口水分有限性 | outlet moisture is finite
    rDenPct : REAL;                  // 分母 (100−w2) | denominator 100 minus w2 [%]
END_VAR
VAR CONSTANT
    DL_DMR_PCT_MAX : REAL := 100.0;  // 含水率上限 | upper moisture limit [%]
    DL_DMR_DEN_MIN : REAL := 1.0E-6; // 除零保护阈值 | division guard threshold [%]
END_VAR

// 段1｜非有限闸（R19）
xFinG := (rFeedKgH = rFeedKgH) AND ((rFeedKgH - rFeedKgH) = 0.0);
xFinW1 := (rMoistInPct = rMoistInPct) AND ((rMoistInPct - rMoistInPct) = 0.0);
xFinW2 := (rMoistOutPct = rMoistOutPct) AND ((rMoistOutPct - rMoistOutPct) = 0.0);
IF (NOT xFinG) OR (NOT xFinW1) OR (NOT xFinW2) THEN
    rWaterRemovedKgH := 0.0;         // 安全值：去水 0 | safe value, zero removal
    rDryMatterKgH := 0.0;
    xReverseMoist := FALSE;
    xValid := FALSE;
    FC_DL_DryerMoistureRemovalCalc := FALSE;
    RETURN;
END_IF

// 段2｜域闸：流量非负、含水率范围、出口含水率不得达 100 %
IF (rFeedKgH < 0.0) OR (rMoistInPct < 0.0) OR (rMoistInPct >= DL_DMR_PCT_MAX)
   OR (rMoistOutPct < 0.0) OR (rMoistOutPct >= DL_DMR_PCT_MAX) THEN
    rWaterRemovedKgH := 0.0;
    rDryMatterKgH := 0.0;
    xReverseMoist := FALSE;
    xValid := FALSE;
    FC_DL_DryerMoistureRemovalCalc := FALSE;
    RETURN;
END_IF

// 段3｜算法：Gd = G×(100−w1)/100；W = Gd×(w1−w2)/(100−w2)
rDryMatterKgH := rFeedKgH * (DL_DMR_PCT_MAX - rMoistInPct) / DL_DMR_PCT_MAX;
rDenPct := DL_DMR_PCT_MAX - rMoistOutPct;
IF rDenPct > DL_DMR_DEN_MIN THEN
    rWaterRemovedKgH := rDryMatterKgH * (rMoistInPct - rMoistOutPct) / rDenPct;
ELSE
    rWaterRemovedKgH := 0.0;         // 理论不可达（段2已排除），防御性兜底 | unreachable defence
END_IF
IF rWaterRemovedKgH < 0.0 THEN
    xReverseMoist := TRUE;           // 回潮工况：信息级告警，出口按 0 发布 | humidification case, informational
    rWaterRemovedKgH := 0.0;
ELSE
    xReverseMoist := FALSE;
END_IF

// 段4｜出口
xValid := TRUE;
FC_DL_DryerMoistureRemovalCalc := TRUE;
END_FUNCTION

(* ---- FC_DL_DryerSolventLoadCalc.st ---- *)
(*
  DL Factory R83 | FC_DL_DryerSolventLoadCalc
  功能：由耗墨量、溶剂配比与排风量估算干燥箱溶剂负荷浓度并做安全裕度校验。
  开源溯源：无（clean-room 自研，依据公开工艺公式，来源=行业通用公式，许可证=MIT，借鉴点=公式结构）
  规则：R1-R21 全遵守
*)
FUNCTION FC_DL_DryerSolventLoadCalc : REAL
VAR_INPUT
    fInkKgH     : REAL; // 单位时间油墨耗量 [kg/h] / Ink consumption rate [kg/h]
    fSolventPct : REAL; // 油墨中溶剂质量占比（0~100）[%] / Solvent mass fraction [%]
    fAirFlowM3H : REAL; // 干燥箱排风量 [m³/h] / Dryer exhaust air flow [m^3/h]
    fLelGm3     : REAL; // 溶剂爆炸下限浓度 [g/m³] / Lower explosive limit [g/m^3]
    fSafetyPct  : REAL; // 安全裕度（允许占 LEL 比例，0~100）[%] / Safety margin of LEL [%]
END_VAR
VAR_OUTPUT
    fSolventKgH : REAL; // 溶剂挥发速率 [kg/h] / Solvent evaporation rate [kg/h]
    fConcGm3    : REAL; // 排风溶剂浓度 [g/m³] / Solvent concentration in exhaust [g/m^3]
    xSafe       : BOOL; // 安全裕度内（TRUE=可继续生产）/ Within safety margin, TRUE = safe
END_VAR
VAR
    fLimitGm3 : REAL; // 允许浓度上限 [g/m³] / Allowed concentration ceiling [g/m^3]
END_VAR
fSolventKgH := 0.0; fConcGm3 := 0.0; xSafe := FALSE;  // 出口预置，安全侧默认不可继续
// 非有限拦截 + 量纲自检（R20/R21）
IF NOT (fInkKgH > -1.0E30 AND fInkKgH < 1.0E30) OR NOT (fSolventPct > -1.0E30 AND fSolventPct < 1.0E30) OR NOT (fAirFlowM3H > -1.0E30 AND fAirFlowM3H < 1.0E30) OR NOT (fLelGm3 > -1.0E30 AND fLelGm3 < 1.0E30) OR NOT (fSafetyPct > -1.0E30 AND fSafetyPct < 1.0E30) OR fInkKgH < 0.0 OR fLelGm3 <= 0.0 OR fSafetyPct <= 0.0 THEN
    FC_DL_DryerSolventLoadCalc := -1.0; RETURN;   // 哨兵 -1：非有限或量纲越界 / Sentinel -1
END_IF
// 溶剂配比域闸：0~100% 之外钳位
IF fSolventPct < 0.0 THEN
    fSolventPct := 0.0;             // 下限钳位 [%] / Clamp lower bound
ELSIF fSolventPct > 100.0 THEN
    fSolventPct := 100.0;           // 上限钳位 [%] / Clamp upper bound
END_IF
// 溶剂挥发速率：kg/h × 质量占比 = kg/h（量纲保持）
fSolventKgH := fInkKgH * (fSolventPct / 100.0);   // 挥发速率 [kg/h] / Evaporation rate [kg/h]
// 排风量零闸后换算浓度：kg/h × 1000 ÷ (m³/h) = g/m³（R4/R21）
IF ABS(fAirFlowM3H) > 1.0E-9 THEN    // 分母显式零闸 / Explicit denominator zero gate
    fConcGm3 := fSolventKgH * 1000.0 / fAirFlowM3H;  // 排风浓度 [g/m³] / Exhaust concentration
ELSE
    fConcGm3 := 0.0;                 // 无排风时浓度不可算，由 xSafe 拦截 / No airflow, default zero
END_IF
// 安全裕度：允许浓度 = LEL × 裕度比例（g/m³ × 无量纲 = g/m³）
fLimitGm3 := fLelGm3 * (fSafetyPct / 100.0);  // 允许浓度上限 [g/m³] / Allowed ceiling [g/m^3]
IF fAirFlowM3H > 0.0 AND fConcGm3 < fLimitGm3 THEN
    xSafe := TRUE;                   // 浓度低于裕度上限 / Concentration below ceiling
ELSE
    xSafe := FALSE;                  // 无排风或浓度超限 / No airflow or over limit
END_IF
FC_DL_DryerSolventLoadCalc := fConcGm3;   // 返回排风浓度 [g/m³] / Return exhaust concentration
END_FUNCTION

(* ---- FC_DL_DryerSteamDemandCalc.st ---- *)
(*
  DL Factory R84 | FC_DL_DryerSteamDemandCalc
  功能：按蒸发水量与汽化潜热折算烘缸蒸汽耗量及单位汽耗
  开源溯源：无（clean-room 自研，依据公开工艺公式，来源=行业通用公式，许可证=MIT，借鉴点=公式结构）
  规则：R1-R16 全遵守
*)
FUNCTION FC_DL_DryerSteamDemandCalc : REAL
VAR_INPUT
    fEvapRateKgh : REAL := 8000.0; // 蒸发水量 [kg/h] / evaporated water rate [kg/h]
    fLatentKjkg : REAL := 2200.0; // 水汽化潜热 [kJ/kg] / latent heat of vaporisation [kJ/kg]
    fSensKjkg : REAL := 250.0; // 水与纸幅显热当量 [kJ/kg] / sensible heat allowance [kJ/kg]
    fSteamEnthKjkg : REAL := 2100.0; // 蒸汽可用焓降 [kJ/kg] / available steam enthalpy drop [kJ/kg]
    fEff : REAL := 0.85; // 烘缸组热效率（0~1） [-] / dryer thermal efficiency [0,1]
    fPaperTph : REAL := 20.0; // 纸机产量 [t/h] / paper machine output [t/h]
END_VAR
VAR_OUTPUT
    fSpecSteam : REAL; // 单位汽耗 [t 汽/t 纸] / specific steam consumption [t/t]
    fEvapKgh : REAL; // 蒸发水量回显（链路校验） [kg/h] / evaporation echo [kg/h]
    xValid : BOOL; // 计算结果有效标志 [-] / calculation valid flag [-]
END_VAR
VAR
    fHeatKjh : REAL; // 需热量 [kJ/h] / heat demand [kJ/h]
    fSteamKgh : REAL; // 蒸汽耗量 [kg/h] / steam demand [kg/h]
END_VAR

// 段 1｜出口预置（R256）
FC_DL_DryerSteamDemandCalc := -1.0; // 哨兵返回 -1（无效） [-] / sentinel return -1, invalid [-]
fSpecSteam := 0.0; // 单位汽耗预置零 [t/t] / specific steam preset zero [t/t]
fEvapKgh := 0.0; // 蒸发量回显预置零 [kg/h] / evaporation echo preset zero [kg/h]
xValid := FALSE; // 计算完成前不认结果 [-] / unusable before calculation [-]

// 段 2｜非有限拦截 + 域闸（R4/R20）
IF NOT (fEvapRateKgh > -1.0E30 AND fEvapRateKgh < 1.0E30) OR NOT (fLatentKjkg > -1.0E30 AND fLatentKjkg < 1.0E30) OR NOT (fSensKjkg > -1.0E30 AND fSensKjkg < 1.0E30) THEN
    RETURN; // 蒸发量与两项热量任一非有限即拒算 [-] / any non finite evaporation or heat term rejected [-]
END_IF
IF NOT (fSteamEnthKjkg > -1.0E30 AND fSteamEnthKjkg < 1.0E30) OR NOT (fEff > -1.0E30 AND fEff < 1.0E30) OR NOT (fPaperTph > -1.0E30 AND fPaperTph < 1.0E30) THEN
    RETURN; // 焓降/效率/产量任一非有限即拒算 [-] / any non finite enthalpy, efficiency or output rejected [-]
END_IF
IF fEvapRateKgh < 0.0 OR fLatentKjkg < 1.0E-9 OR fSensKjkg < 0.0 THEN
    RETURN; // 蒸发量非负 + 潜热正域闸 [kg/h, kJ/kg] / non negative evaporation and positive latent heat gate [-]
END_IF
IF fSteamEnthKjkg < 1.0E-9 OR fEff < 1.0E-9 OR fPaperTph < 1.0E-9 THEN
    RETURN; // 焓降/效率/产量正域分母闸（防除零） [kJ/kg, t/h] / positive denominator gate [kJ/kg, t/h]
END_IF
IF fEff > 1.0 THEN
    RETURN; // 效率上限闸：大于一违反热力学 [-] / efficiency above one is not physical [-]
END_IF

// 段 3｜需热量与蒸汽耗量
fHeatKjh := fEvapRateKgh * (fLatentKjkg + fSensKjkg); // kg/h × kJ/kg = kJ/h / [kg/h] × [kJ/kg] = [kJ/h]
fSteamKgh := (fHeatKjh / fSteamEnthKjkg) / fEff; // kJ/h ÷ kJ/kg = kg/h；÷ 无量纲 仍 kg/h / [kJ/h] / [kJ/kg] / [-] = [kg/h]
IF NOT (fSteamKgh > -1.0E30 AND fSteamKgh < 1.0E30) THEN
    RETURN; // 结果非有限再拦一次 [-] / second finiteness gate [-]
END_IF

// 段 4｜单位汽耗 = 汽量 / 纸量（同除 kg/h 得无量纲，即 t/t）
fSpecSteam := fSteamKgh / (fPaperTph * 1000.0); // kg/h ÷ (t/h × 1000 kg/t) = 无量纲（t 汽/t 纸） / [kg/h] / [kg/h] = [-] = [t/t]
IF NOT (fSpecSteam > -1.0E30 AND fSpecSteam < 1.0E30) THEN
    RETURN; // 结果非有限再拦一次 [-] / second finiteness gate [-]
END_IF
fEvapKgh := fEvapRateKgh; // 回显蒸发水量 [kg/h] / echo the evaporated water [kg/h]
xValid := TRUE; // 链路有效 [-] / chain valid [-]
FC_DL_DryerSteamDemandCalc := fSteamKgh; // 返回蒸汽耗量 [kg/h] / return the steam demand [kg/h]
END_FUNCTION

(* ---- FC_DL_DyeExhaustionCalc.st ---- *)
(*
  Name: FC_DL_DyeExhaustionCalc
  Category: DL_Process
  Version: 1.0.0
  Round: R91 / 2026-11-25
  开源溯源：clean-room 自研（族 间歇式溢流染色与丝光整理，ST 开源生态实测 0 命中，无外部代码引入）
  功能：1) 上染率（竭染率）按「初始与残液浓度差」计算：
           E = (C0 − C1) / C0 * 100，C0 为初始染浴浓度、C1 为残液（或染后液）浓度，
           两者取同一稀释倍数下的分光光度换算值，故可直接相减；
           分母固定为初始浓度（上染率是「初始染料中被纤维吸收的比例」）。
        2) 派生量：fUptakeGpl 为单位液量被纤维吸收的染料量 [g/L]，
           用于核算染化料成本与残液回用价值。
        3) 双向异常判定：E < 0（残液比初始还浓，说明浓度测量错位或补料干扰）判 xNegative；
           E > 100（吸收量超过投加量，违反质量守恒）判 xOverHundred。
           两者任一成立即判无效，绝不把异常值当作合格上染率。
  边界条件：1) 非有限值闸：两路实值入参先过 NOT(x > -DL_BIG AND x < DL_BIG)，同时拦 NaN 与 Inf，
           命中即闸断实值通路（上染率与吸收量强制 0.0 且置负向异常位，保守侧），不得只置标志（R19）。
        2) 初始浓度零闸：fInitConcGpl 必须 > DL_EPS（上染率式的分母），
           为零则结果发散，判无效并清零，绝不输出「无穷大上染率」。
        3) 浓度非负闸：残液浓度不得为负（负浓度属分光光度计基线漂移或比色皿污染），判无效。
        4) 判据取原始值（R24）：双向异常判定使用钳制前的 _fExhaustRawPct，钳制只作用于输出。
        5) 物理域钳制：上染率钳 0.0 ~ DL_PCT_HI；吸收量钳 0.0 ~ 初始浓度（吸收不可能超过投加）。
        6) 纯函数无状态：上染率的实时趋势与「终点判定」（达 95 % 即转水洗）由上层染缸序 FB 承担。
  量纲自证：E = (g/L − g/L) / (g/L) * 100 = 无因次百分数 [%]；
           fUptakeGpl = (g/L) − (g/L) = g/L，减法两侧同量纲，量纲合法。
  修订历史 Revision :
    2026-11-25  v1.0.0  R91 首版
*)

FUNCTION FC_DL_DyeExhaustionCalc : BOOL
VAR_INPUT
    fInitConcGpl     : REAL;   // 初始染浴染料浓度 [g/L] / Initial dye bath concentration [g/L]
    fResidualConcGpl : REAL;   // 残液染料浓度 [g/L] / Residual dye concentration [g/L]
END_VAR
VAR_OUTPUT
    fExhaustPct      : REAL;   // 上染率（竭染率）[%] / Dye exhaustion [%]
    fUptakeGpl       : REAL;   // 单位液量被吸收的染料量 [g/L] / Dye taken up per litre of bath [g/L]
    xNegative        : BOOL;   // 上染率为负（方向异常）标志 [bool] / Negative exhaustion flag [bool]
    xOverHundred     : BOOL;   // 上染率超 100 %（违反守恒）标志 [bool] / Exhaustion over 100 percent flag [bool]
    xValid           : BOOL;   // 计算有效标志 [bool] / Calculation valid flag [bool]
END_VAR
VAR
    _fUptakeRawGpl   : REAL;   // 钳制前的吸收量 [g/L] / Raw uptake before limiting [g/L]
    _fExhaustRawPct  : REAL;   // 钳制前的原始上染率 [%] / Raw exhaustion before limiting [%]
END_VAR
VAR CONSTANT
    DL_EPS           : REAL := 1.0E-9;    // 数值零闸阈值 [-] / Numeric zero gate threshold [-]
    DL_BIG           : REAL := 1.0E12;    // 非有限值闸量级上限 [-] / Finiteness gate magnitude [-]
    DL_PCT           : REAL := 100.0;     // 百分比换算因子 [%] / Percent conversion factor [%]
    DL_CONC_HI_GPL   : REAL := 200.0;     // 染料浓度量级闸上限 [g/L] / Concentration magnitude upper bound [g/L]
END_VAR

(* —— 段 1：非有限值闸（R19：闸断实值通路；失效侧置负向异常，保守侧） —— *)
IF NOT (fInitConcGpl > -DL_BIG AND fInitConcGpl < DL_BIG)
   OR NOT (fResidualConcGpl > -DL_BIG AND fResidualConcGpl < DL_BIG) THEN
    fExhaustPct := 0.0;                     // 输出强制 0.0，切断污染源 / Force zero, cut polluted path
    fUptakeGpl := 0.0;                      // 吸收量强制 0.0 / Uptake forced to zero
    xNegative := TRUE;                      // 失效侧按方向异常处理 / Treat as abnormal when invalid
    xOverHundred := FALSE;                  // 失效侧超百位保持假 / Over-hundred stays false
    xValid := FALSE;                        // 有效位清零 / Validity cleared
    FC_DL_DyeExhaustionCalc := FALSE;       // 返回码与有效位同源 / Return mirrors validity
    RETURN;                                 // 立即退出 / Immediate exit
END_IF

(* —— 段 2：初始浓度零闸与量级闸（分母为初始浓度） —— *)
IF (fInitConcGpl <= DL_EPS)                                       // 初始浓度不可为零
   OR (fResidualConcGpl < 0.0)                                    // 残液浓度不得为负
   OR (fInitConcGpl > DL_CONC_HI_GPL)                             // 初始浓度量级闸
   OR (fResidualConcGpl > DL_CONC_HI_GPL) THEN                    // 残液浓度量级闸
    fExhaustPct := 0.0;                     // 分母为零即不可算 / No denominator, no ratio
    fUptakeGpl := 0.0;                      // 吸收量不可算 / Uptake not computable
    xNegative := TRUE;                      // 按方向异常处理（保守侧）/ Treat as abnormal
    xOverHundred := FALSE;                  // 超百位保持假 / Over-hundred stays false
    xValid := FALSE;                        // 判无效 / Invalid
    FC_DL_DyeExhaustionCalc := FALSE;       // 返回码同步 / Return synchronised
    RETURN;                                 // 提前退出 / Early exit
END_IF

(* —— 段 3：主算式（不钳制，先出原始值供段 4 判据使用，R24） —— *)
_fUptakeRawGpl := fInitConcGpl - fResidualConcGpl;                                // 吸收量 [g/L]
_fExhaustRawPct := _fUptakeRawGpl / fInitConcGpl * DL_PCT;                        // 上染率 [%]

(* —— 段 4：判据（取原始值；单点 BOOL 聚合避免多处赋 FALSE 覆盖） —— *)
xNegative := (_fExhaustRawPct < 0.0);                                             // 残液比初始还浓：方向异常
xOverHundred := (_fExhaustRawPct > DL_PCT);                                       // 超 100 %：违反质量守恒
xValid := (NOT xNegative) AND (NOT xOverHundred)                                  // 双向异常位均不成立
          AND (_fUptakeRawGpl >= 0.0);                                            // 吸收量不得为负

(* —— 段 5：输出单点写盘（钳制到物理域内，判定结果已在段 4 定案） —— *)
fExhaustPct := LIMIT(0.0, _fExhaustRawPct, DL_PCT);                               // 上染率钳 0..100 [%]
fUptakeGpl := LIMIT(0.0, _fUptakeRawGpl, fInitConcGpl);                            // 吸收量钳 0..初始浓度 [g/L]
FC_DL_DyeExhaustionCalc := xValid;                                                // 返回码：TRUE = 计算可信

END_FUNCTION

(* ---- FC_DL_DyeLiquorRatioCalc.st ---- *)
(*
  DL Factory R83 | FC_DL_DyeLiquorRatioCalc
  功能：按织物重量与浴比算染浴总液量，并给出需补加液量与补加耗时。
  开源溯源：无（clean-room 自研，依据公开工艺公式，来源=行业通用公式，许可证=MIT，借鉴点=公式结构）
  规则：R1-R21 全遵守
*)
FUNCTION FC_DL_DyeLiquorRatioCalc : REAL
VAR_INPUT
    fFabricKg    : REAL; // 投染织物重量 [kg] / Fabric batch weight [kg]
    fLiquorRatio : REAL; // 浴比（每 kg 织物配液量）[L/kg] / Liquor ratio [L/kg]
    fBathVolL    : REAL; // 染缸现有液量 [L] / Existing bath volume [L]
    fAddRateLpm  : REAL; // 补水/补液流量 [L/min] / Replenish flow rate [L/min]
END_VAR
VAR_OUTPUT
    fTotalL : REAL; // 工艺要求总液量 [L] / Required total liquor volume [L]
    fAddL   : REAL; // 尚需补加液量（负偏差按零）[L] / Volume still to add, clamped at zero [L]
    fAddMin : REAL; // 补加所需时间 [min] / Time needed to add [min]
    xValid  : BOOL; // 计算有效性标志 / Calculation validity flag
END_VAR
VAR
    fDiffL : REAL; // 总液量与现有液量之差 [L] / Volume difference [L]
END_VAR
fTotalL := 0.0; fAddL := 0.0; fAddMin := 0.0; xValid := FALSE;  // 出口预置（R256）
// 非有限拦截 + 量纲自检（R20/R21）
IF NOT (fFabricKg > -1.0E30 AND fFabricKg < 1.0E30) OR NOT (fLiquorRatio > -1.0E30 AND fLiquorRatio < 1.0E30) OR NOT (fBathVolL > -1.0E30 AND fBathVolL < 1.0E30) OR NOT (fAddRateLpm > -1.0E30 AND fAddRateLpm < 1.0E30) OR fFabricKg <= 0.0 OR fLiquorRatio <= 0.0 OR fBathVolL < 0.0 THEN
    FC_DL_DyeLiquorRatioCalc := -1.0; RETURN;   // 哨兵 -1：非有限或量纲越界 / Sentinel -1
END_IF
// 浴比域闸：0.5~50 L/kg 之外钳位（工艺可执行区间）
IF fLiquorRatio < 0.5 THEN
    fLiquorRatio := 0.5;            // 下限钳位 [L/kg] / Clamp to 0.5 L/kg
ELSIF fLiquorRatio > 50.0 THEN
    fLiquorRatio := 50.0;           // 上限钳位 [L/kg] / Clamp to 50 L/kg
END_IF
// 总液量：kg × L/kg = L（量纲自洽，kg 约去）
fTotalL := fFabricKg * fLiquorRatio;   // 工艺总液量 [L] / Required total volume [L]
// 补加量：差值负值按零，避免抽液反算（单向补加语义）
fDiffL := fTotalL - fBathVolL;      // 液量差 [L] / Volume difference [L]
IF fDiffL > 0.0 THEN
    fAddL := fDiffL;                // 需要补加 [L] / Volume to add [L]
ELSE
    fAddL := 0.0;                   // 已够量，不抽液 [L] / Already sufficient [L]
END_IF
// 补加时间：L ÷ (L/min) = min，流量分母显式零闸（R4/R21）
IF ABS(fAddRateLpm) > 1.0E-9 THEN   // 分母显式零闸 / Explicit denominator zero gate
    fAddMin := fAddL / fAddRateLpm; // 补加时间 [min] / Add time [min]
ELSE
    fAddMin := 0.0;                 // 无流量时不可估时，缺省零 / No flow, default zero
END_IF
xValid := TRUE; FC_DL_DyeLiquorRatioCalc := fTotalL;  // 链路有效并返回总液量 [L] / Return volume
END_FUNCTION

(* ---- FC_DL_DyeShadeDeltaCalc.st ---- *)
(*
  Name: FC_DL_DyeShadeDeltaCalc
  Category: DL_Process
  Version: 1.0.0
  Round: R91 / 2026-11-25
  开源溯源：clean-room 自研（族 间歇式溢流染色与丝光整理，ST 开源生态实测 0 命中，无外部代码引入）
  功能：1) 色差按 CIE76 色差公式（CIE 1976 L*a*b* 空间的欧氏距离）计算：
           dE = SQRT(dL^2 + da^2 + db^2)，
           其中 dL = L_sample − L_std、da = a_sample − a_std、db = b_sample − b_std，
           标准样与被测样必须取自同一光源/观察者条件（D65 / 10 deg）下的测色值。
           CIE76 为不带权重的等距公式，计算稳定、可复现，是染厂判色的基准口径。
        2) 三档判定（nGrade）：0 = 合格（dE <= fPassDE）、1 = 返修（可回修，<= fReworkDE）、
           2 = 回修（超出返修上限，须改色或降级），两级阈值由工艺按订单要求给定。
        3) 亮度分量 dL 单独输出：dL 与 |da|/|db| 的大小关系决定纠偏方向
           （dL 主导调深浅，a/b 主导调色光），供配色系统选配方。
  边界条件：1) 非有限值闸：六路 Lab 入参与两路阈值先过 NOT(x > -DL_BIG AND x < DL_BIG)，
           同时拦 NaN 与 Inf，命中即闸断实值通路（色差强制 0.0 且分级置 2 = 回修，保守侧），
           不得只置标志（R19）。
        2) 量级闸：Lab 各分量必须落在 [-DL_LAB_SPAN, +DL_LAB_SPAN] 内（L* 为 0~100、a*/b* 约 ±128），
           越域说明色差仪标定丢失或数据通道错位，判无效。
        3) 阈值域闸：须满足 0.0 < fPassDE < fReworkDE，且 fReworkDE <= DL_DE_HI，
           否则三档判定区间为空、某档永不触发，判无效并把分级置 2（保守侧）。
        4) 平方和防溢出：三个分量的平方和先做量级闸（各分量有界 => 平方和有界），
           SQRT 前不再额外钳制，量级闸是唯一入口，避免「先钳后判」使判据恒真（R24）。
        5) 判据取原始值（R24）：三档判定使用未钳制的 _fDeltaERaw，钳制只作用于输出数值。
        6) 纯函数无状态：多测点平均色差与首件/末件比对由上层判色模块承担。
  量纲自证：dL / da / db 与 Lab 分量同为无因次色度值（CIE L*a*b* 为无量纲量）；
           dE = SQRT(无因次^2 * 3) = 无因次，与阈值 fPassDE / fReworkDE 同量纲。
  修订历史 Revision :
    2026-11-25  v1.0.0  R91 首版
*)

FUNCTION FC_DL_DyeShadeDeltaCalc : BOOL
VAR_INPUT
    fLStd            : REAL;   // 标准样明度 L* [-]/ Standard lightness L* [-]
    fAStd            : REAL;   // 标准样红绿色度 a* [-]/ Standard redness-greenness a* [-]
    fBStd            : REAL;   // 标准样黄蓝色度 b* [-]/ Standard yellowness-blueness b* [-]
    fLSample         : REAL;   // 被测样明度 L* [-]/ Sample lightness L* [-]
    fASample         : REAL;   // 被测样红绿色度 a* [-]/ Sample redness-greenness a* [-]
    fBSample         : REAL;   // 被测样黄蓝色度 b* [-]/ Sample yellowness-blueness b* [-]
    fPassDE          : REAL;   // 合格色差上限 [-]/ Colour difference acceptance limit [-]
    fReworkDE        : REAL;   // 返修色差上限 [-]/ Colour difference rework limit [-]
END_VAR
VAR_OUTPUT
    fDeltaE          : REAL;   // 色差 dE（CIE76）[-]/ Colour difference dE, CIE76 [-]
    fDeltaL          : REAL;   // 明度差 dL（带符号）[-]/ Lightness difference, signed [-]
    nGrade           : INT;    // 判定 0=合格 1=返修 2=回修 [level] / Verdict 0=pass 1=reworkable 2=reject [level]
    xValid           : BOOL;   // 计算有效标志 [bool] / Calculation valid flag [bool]
END_VAR
VAR
    _fDeltaL         : REAL;   // 明度差分量 [-]/ Lightness difference component [-]
    _fDeltaA         : REAL;   // 红绿色度差分量 [-]/ Redness-greenness difference component [-]
    _fDeltaB         : REAL;   // 黄蓝色度差分量 [-]/ Yellowness-blueness difference component [-]
    _fSumSq          : REAL;   // 三分量平方和 [-]/ Sum of squared components [-]
    _fDeltaERaw      : REAL;   // 未钳制的色差 [-]/ Unclamped colour difference [-]
END_VAR
VAR CONSTANT
    DL_BIG           : REAL := 1.0E12;    // 非有限值闸量级上限 [-] / Finiteness gate magnitude [-]
    DL_EPS           : REAL := 1.0E-9;    // 数值零闸阈值 [-] / Numeric zero gate threshold [-]
    DL_LAB_SPAN      : REAL := 500.0;     // Lab 分量量级闸跨度 [-] / Lab component magnitude gate span [-]
    DL_DE_HI         : REAL := 500.0;     // 色差物理上限 [-] / Colour difference physical upper bound [-]
    DL_GRADE_OK      : INT := 0;          // 判定：合格 [level] / Verdict: pass [level]
    DL_GRADE_REWORK  : INT := 1;          // 判定：返修 [level] / Verdict: reworkable [level]
    DL_GRADE_REJECT  : INT := 2;          // 判定：回修 [level] / Verdict: reject [level]
END_VAR

(* —— 段 1：非有限值闸（R19：闸断实值通路；失效侧分级置回修） —— *)
IF NOT (fLStd > -DL_BIG AND fLStd < DL_BIG)
   OR NOT (fAStd > -DL_BIG AND fAStd < DL_BIG)
   OR NOT (fBStd > -DL_BIG AND fBStd < DL_BIG)
   OR NOT (fLSample > -DL_BIG AND fLSample < DL_BIG)
   OR NOT (fASample > -DL_BIG AND fASample < DL_BIG)
   OR NOT (fBSample > -DL_BIG AND fBSample < DL_BIG)
   OR NOT (fPassDE > -DL_BIG AND fPassDE < DL_BIG)
   OR NOT (fReworkDE > -DL_BIG AND fReworkDE < DL_BIG) THEN
    fDeltaE := 0.0;                         // 输出强制 0.0，切断污染源 / Force zero, cut polluted path
    fDeltaL := 0.0;                         // 明度差强制 0.0 / Lightness difference forced to zero
    nGrade := DL_GRADE_REJECT;              // 失效侧按回修处理（保守侧）/ Treat as reject when invalid
    xValid := FALSE;                        // 有效位清零 / Validity cleared
    FC_DL_DyeShadeDeltaCalc := FALSE;       // 返回码与有效位同源 / Return mirrors validity
    RETURN;                                 // 立即退出 / Immediate exit
END_IF

(* —— 段 2：量级闸与阈值域闸（Lab 越域与阈值倒置都使判定失效） —— *)
IF (ABS(fLStd) > DL_LAB_SPAN) OR (ABS(fAStd) > DL_LAB_SPAN) OR (ABS(fBStd) > DL_LAB_SPAN)
   OR (ABS(fLSample) > DL_LAB_SPAN) OR (ABS(fASample) > DL_LAB_SPAN) OR (ABS(fBSample) > DL_LAB_SPAN)
   OR (fPassDE <= 0.0) OR (fReworkDE <= fPassDE) OR (fReworkDE > DL_DE_HI) THEN
    fDeltaE := 0.0;                         // 量级越域即不可算 / Out of range, not computable
    fDeltaL := 0.0;                         // 明度差不可算 / Lightness difference not computable
    nGrade := DL_GRADE_REJECT;              // 按回修处理（保守侧）/ Treat as reject
    xValid := FALSE;                        // 判无效 / Invalid
    FC_DL_DyeShadeDeltaCalc := FALSE;       // 返回码同步 / Return synchronised
    RETURN;                                 // 提前退出 / Early exit
END_IF

(* —— 段 3：主算式（CIE76 欧氏距离；分量已由段 2 保证有界，平方和不会溢出） —— *)
_fDeltaL := fLSample - fLStd;                                                     // 明度差 [-]
_fDeltaA := fASample - fAStd;                                                     // 红绿色度差 [-]
_fDeltaB := fBSample - fBStd;                                                     // 黄蓝色度差 [-]
_fSumSq := _fDeltaL * _fDeltaL + _fDeltaA * _fDeltaA + _fDeltaB * _fDeltaB;       // 平方和 [-]
_fDeltaERaw := SQRT(_fSumSq);                                                     // 色差 [-]
fDeltaL := _fDeltaL;                                                              // 明度差出口（供纠偏方向）

(* —— 段 4：三档判定（取原始色差；由上到下判，区间互斥且完整） —— *)
IF _fDeltaERaw <= fPassDE THEN
    nGrade := DL_GRADE_OK;                  // 合格
ELSIF _fDeltaERaw <= fReworkDE THEN
    nGrade := DL_GRADE_REWORK;              // 可返修
ELSE
    nGrade := DL_GRADE_REJECT;              // 回修/降级
END_IF

xValid := (_fDeltaERaw >= 0.0)                                                    // 色差恒非负（SQRT 性质）
          AND (_fDeltaERaw <= DL_DE_HI);                                          // 不超物理上限（量级异常）

(* —— 段 5：输出单点写盘（钳制到物理域内，判定结果已在段 4 定案） —— *)
fDeltaE := LIMIT(0.0, _fDeltaERaw, DL_DE_HI);                                     // 色差钳物理域 [-]
FC_DL_DyeShadeDeltaCalc := xValid;                                                // 返回码：TRUE = 计算可信

END_FUNCTION

(* ---- FC_DL_ElectrodeCompactionRatioCalc.st ---- *)
(*
  Name: FC_DL_ElectrodeCompactionRatioCalc
  Category: DL_Process
  Version: 1.0.0
  Round: R90 / 2026-11-25
  开源溯源：clean-room 自研（族 锂电极片涂布辊压，ST 开源生态实测 0 命中，无外部代码引入）
  功能：1) 压实比按「辊压后密度 / 辊压前（来料）密度」计算，是无因次的密实化倍数。
           该比值与面密度、厚度无关，只反映辊压工序本身的密实效果，适合作为辊压工艺窗口判据。
        2) 工艺窗口判定 xInWindow：压实比落在 [fRatioMin, fRatioMax] 闭区间内即判合格。
           窗口上下限由组态给出，本件不硬编码工艺值；上下限本身做合法性校验（下限须 > 1，
           因为压实比 = 1 表示完全未压实，< 1 表示减薄的反向过程，均不属辊压工艺窗口）。
  边界条件：1) 非有限值闸：四路实值入参统一过 NOT(x > -DL_BIG AND x < DL_BIG)，
           同时拦 NaN 与 Inf，命中即拦断实值通路（fRatio 强制 0.0、xInWindow 强制 FALSE）并置无效（R19），
           无效数据不得判合格。
        2) 分母零闸：ABS(fGreenGcm3) > DL_EPS 才允许相除（来料密度为 0 时比值无定义）。
        3) 负值闸：两个密度任一为负、窗口上下限任一为负均判无效。
        4) 窗口组态闸：fRatioMax 必须 >= fRatioMin，否则窗口为空集、合格判据恒假（组态错误）；
           fRatioMin 必须 >= 1.0，否则窗口包含「未压实或减薄」的非物理区间。
        5) 饱和钳制：压实比钳 0 ~ DL_RATIO_MAX(20)，防极小来料密度把比值放大到无意义量级。
  量纲自证：fRatio = (g/cm3) / (g/cm3) = 无因次 [-]；
           窗口上下限同为无因次，与 fRatio 同量纲后方可比较；本件无跨量纲相加。
*)

FUNCTION FC_DL_ElectrodeCompactionRatioCalc : BOOL
VAR_INPUT
    fCompactionGcm3 : REAL;   // 辊压后压实密度 [g/cm3] / Post-calendering compaction density [g/cm3]
    fGreenGcm3      : REAL;   // 辊压前来料密度 [g/cm3] / Incoming green density [g/cm3]
    fRatioMin       : REAL;   // 工艺窗口下限 [-] / Process window lower limit [-]
    fRatioMax       : REAL;   // 工艺窗口上限 [-] / Process window upper limit [-]
END_VAR
VAR_OUTPUT
    fRatio          : REAL;   // 压实比 [-] / Compaction ratio [-]
    xInWindow       : BOOL;   // 落在工艺窗口内 [bool] / Inside process window flag [bool]
    xValid          : BOOL;   // 计算有效标志 [bool] / Calculation valid flag [bool]
END_VAR
VAR
    _fRatioRaw      : REAL;   // 未饱和的压实比 [-] / Raw compaction ratio [-]
END_VAR
VAR CONSTANT
    DL_EPS          : REAL := 1.0E-9;    // 分母零闸阈值 [-] / Division-zero gate threshold [-]
    DL_BIG          : REAL := 1.0E12;    // 非有限值闸量级上限 [-] / Finiteness gate magnitude [-]
    DL_RATIO_MAX    : REAL := 20.0;      // 压实比饱和上限 [-] / Compaction ratio saturation ceiling [-]
    DL_RATIO_MIN_OK : REAL := 1.0;       // 压实比物理下限（未压实）[-] / Physical lower bound [-]
END_VAR

(* —— 段 1：非有限值闸（R19：四路入参全覆盖，拦 NaN 与 Inf） —— *)
IF NOT (fCompactionGcm3 > -DL_BIG AND fCompactionGcm3 < DL_BIG)
   OR NOT (fGreenGcm3 > -DL_BIG AND fGreenGcm3 < DL_BIG)
   OR NOT (fRatioMin > -DL_BIG AND fRatioMin < DL_BIG)
   OR NOT (fRatioMax > -DL_BIG AND fRatioMax < DL_BIG) THEN
    fRatio := 0.0;                          // 输出强制 0.0 / Output forced to zero
    xInWindow := FALSE;                     // 窗口标志强制 FALSE / Window flag forced off
    xValid := FALSE;                        // 有效位清零 / Validity cleared
    FC_DL_ElectrodeCompactionRatioCalc := FALSE;   // 返回码同源 / Return mirrors validity
    RETURN;                                 // 立即退出 / Immediate exit
END_IF

(* —— 段 2：分母零闸（R4：来料密度是比值分母） —— *)
IF ABS(fGreenGcm3) <= DL_EPS THEN
    fRatio := 0.0;                          // 输出强制 0.0 / Output forced to zero
    xInWindow := FALSE;                     // 窗口标志强制 FALSE / Window flag forced off
    xValid := FALSE;                        // 判无效 / Invalid
    FC_DL_ElectrodeCompactionRatioCalc := FALSE;   // 返回码同步 / Return synchronised
    RETURN;                                 // 提前退出 / Early exit
END_IF

(* —— 段 3：负值闸（密度与窗口限值均不可为负） —— *)
IF (fCompactionGcm3 < 0.0) OR (fGreenGcm3 < 0.0) OR (fRatioMin < 0.0) OR (fRatioMax < 0.0) THEN
    fRatio := 0.0;                          // 输出强制 0.0 / Output forced to zero
    xInWindow := FALSE;                     // 窗口标志强制 FALSE / Window flag forced off
    xValid := FALSE;                        // 判无效 / Invalid
    FC_DL_ElectrodeCompactionRatioCalc := FALSE;   // 返回码同步 / Return synchronised
    RETURN;                                 // 提前退出 / Early exit
END_IF

(* —— 段 4：主算式（R22 方向自核：压实后密度在分子、来料密度在分母，比值必 >= 1） —— *)
_fRatioRaw := fCompactionGcm3 / fGreenGcm3;                       // 压实比 [-]

(* —— 段 5：输出单点写盘（饱和钳制后判窗口，保证判据与出口同源） —— *)
fRatio := LIMIT(0.0, _fRatioRaw, DL_RATIO_MAX);                   // 压实比 [-]

(* —— 段 6：有效位单点聚合（窗口组态合法性 + 密度为正） —— *)
xValid := (fGreenGcm3 > DL_EPS)                                   // 来料密度为正
          AND (fCompactionGcm3 > DL_EPS)                          // 压实密度为正
          AND (fRatioMax >= fRatioMin)                            // 窗口非空
          AND (fRatioMin >= DL_RATIO_MIN_OK);                     // 下限不落入非物理区间

(* —— 段 7：工艺窗口判定（闭区间，边界值算合格） —— *)
xInWindow := xValid AND (fRatio >= fRatioMin) AND (fRatio <= fRatioMax);
FC_DL_ElectrodeCompactionRatioCalc := xValid;                     // 返回码：TRUE = 计算可信

END_FUNCTION

(* ---- FC_DL_ElectrodePorosityCalc.st ---- *)
(*
  Name: FC_DL_ElectrodePorosityCalc
  Category: DL_Process
  Version: 1.0.0
  Round: R90 / 2026-11-25
  开源溯源：clean-room 自研（族 锂电极片涂布辊压，ST 开源生态实测 0 命中，无外部代码引入）
  功能：1) 极片孔隙率按「孔隙体积占表观体积的比例」计算。表观体积 V = 涂层质量 / 压实密度，
           固体实体体积 V_s = 涂层质量 / 真密度，孔隙体积 = V − V_s，
           故孔隙率 = 1 − 压实密度 / 真密度，乘 100 转百分数。
           该式与涂层质量无关（质量在比值中消去），只取决于两个密度之比。
        2) 用于辊压工序的压实程度评价：孔隙率过低会导致电解液浸润困难与析锂风险，
           过高则电子导电网络接触不良、能量密度不足，故需落在工艺窗口内。
  边界条件：1) 非有限值闸：两路实值入参统一过 NOT(x > -DL_BIG AND x < DL_BIG)，
           同时拦 NaN 与 Inf，命中即拦断实值通路（fPorosityPct 强制 0.0）并置无效（R19）。
        2) 分母零闸：ABS(fTrueDensityGcm3) > DL_EPS 才允许相除（真密度为 0 无物理意义）。
        3) 负值闸：两个密度任一为负判无效（不取绝对值掩盖反向）。
        4) 物理域校验：压实密度必须严格小于真密度，否则孔隙率为负（固体体积大于表观体积，
           不可能），判无效且输出钳 0；结果同时钳到 0 ~ 100 % 的物理域。
        5) 量程校验：真密度钳 0 ~ DL_RHO_MAX(10 g/cm3)、压实密度同域，越域钳边界算参考值但置无效；
           真密度为 0 与「三元材料 2.0~5.0 g/cm3」的实际量程差距过大，故另设 DL_RHO_MIN(0.5 g/cm3)
           作为可信下限，低于该值视为组态或传感器异常。
  量纲自证：孔隙率 = 1 − (g/cm3) / (g/cm3) = 1 − 无因次 = 无因次，乘 100 得 [%]；
           密度比无量纲，厚度/质量/体积项均已通过密度定义消去，无跨量纲相加。
*)

FUNCTION FC_DL_ElectrodePorosityCalc : BOOL
VAR_INPUT
    fCompactionGcm3  : REAL;   // 极片压实密度 [g/cm3] / Electrode compaction density [g/cm3]
    fTrueDensityGcm3 : REAL;   // 材料真密度 [g/cm3] / Material true density [g/cm3]
END_VAR
VAR_OUTPUT
    fPorosityPct     : REAL;   // 极片孔隙率 [%] / Electrode porosity [%]
    xValid           : BOOL;   // 计算有效标志 [bool] / Calculation valid flag [bool]
END_VAR
VAR
    _fDensityRatio   : REAL;   // 压实密度 / 真密度 [-] / Compaction to true density ratio [-]
    _fPorosityRawPct : REAL;   // 未饱和的孔隙率 [%] / Raw porosity [%]
END_VAR
VAR CONSTANT
    DL_EPS           : REAL := 1.0E-9;    // 分母零闸阈值 [-] / Division-zero gate threshold [-]
    DL_BIG           : REAL := 1.0E12;    // 非有限值闸量级上限 [-] / Finiteness gate magnitude [-]
    DL_PCT           : REAL := 100.0;     // 百分比换算因子 [%] / Percent conversion factor [%]
    DL_RHO_MIN       : REAL := 0.50;      // 密度可信下限 [g/cm3] / Density credibility low [g/cm3]
    DL_RHO_MAX       : REAL := 10.0;      // 密度量程上限 [g/cm3] / Density range ceiling [g/cm3]
END_VAR

(* —— 段 1：非有限值闸（R19：闸断实值通路，NaN 不得进入比值） —— *)
IF NOT (fCompactionGcm3 > -DL_BIG AND fCompactionGcm3 < DL_BIG)
   OR NOT (fTrueDensityGcm3 > -DL_BIG AND fTrueDensityGcm3 < DL_BIG) THEN
    fPorosityPct := 0.0;                    // 输出强制 0.0 / Output forced to zero
    xValid := FALSE;                        // 有效位清零 / Validity cleared
    FC_DL_ElectrodePorosityCalc := FALSE;   // 返回码同源 / Return mirrors validity
    RETURN;                                 // 立即退出 / Immediate exit
END_IF

(* —— 段 2：分母零闸（R4：真密度是比值分母） —— *)
IF ABS(fTrueDensityGcm3) <= DL_EPS THEN
    fPorosityPct := 0.0;                    // 输出强制 0.0 / Output forced to zero
    xValid := FALSE;                        // 判无效 / Invalid
    FC_DL_ElectrodePorosityCalc := FALSE;   // 返回码同步 / Return synchronised
    RETURN;                                 // 提前退出 / Early exit
END_IF

(* —— 段 3：负值闸（密度为负无物理意义，不取绝对值掩盖） —— *)
IF (fCompactionGcm3 < 0.0) OR (fTrueDensityGcm3 < 0.0) THEN
    fPorosityPct := 0.0;                    // 输出强制 0.0 / Output forced to zero
    xValid := FALSE;                        // 判无效 / Invalid
    FC_DL_ElectrodePorosityCalc := FALSE;   // 返回码同步 / Return synchronised
    RETURN;                                 // 提前退出 / Early exit
END_IF

(* —— 段 4：主算式（R22 方向自核：压实密度在分子，真密度在分母，二者不可交换） —— *)
_fDensityRatio := fCompactionGcm3 / fTrueDensityGcm3;             // 密度比 [-]
_fPorosityRawPct := (1.0 - _fDensityRatio) * DL_PCT;              // 孔隙率 [%]

(* —— 段 5：输出单点写盘（钳到 0~100 % 物理域，负孔隙率不得流出） —— *)
fPorosityPct := LIMIT(0.0, _fPorosityRawPct, DL_PCT);             // 孔隙率 [%]

(* —— 段 6：有效位单点聚合（物理域 + 密度量程） —— *)
xValid := (fCompactionGcm3 < fTrueDensityGcm3)                    // 压实密度必须小于真密度
          AND (fTrueDensityGcm3 >= DL_RHO_MIN)                    // 真密度不低于可信下限
          AND (fTrueDensityGcm3 <= DL_RHO_MAX)                    // 真密度不越量程
          AND (fCompactionGcm3 <= DL_RHO_MAX);                    // 压实密度不越量程
FC_DL_ElectrodePorosityCalc := xValid;                            // 返回码：TRUE = 计算可信

END_FUNCTION

(* ---- FC_DL_ExtrusionBilletHeatCalc.st ---- *)
(*
  Component : FC_DL_ExtrusionBilletHeatCalc
  Category  : DL_Process
  Type      : FC
  Complexity: C2
  VERSION   : v1.0.0
  功能      : 铝挤压铸锭感应加热负荷核算：按锭重/比热/温升/效率算所需电功率与总能耗 kWh。
  开源溯源  : 道莅原创 clean-room 自研（无外部代码引用）｜License: MIT
  边界条件  : ① 锭重、加热时长须 > 1e-9，锭数须 >= 1，效率须在 (0, 100] % 内，否则返回哨兵 -1；
              ② 温升目标不高于起始温度时，能耗与功率均输出 0 且 xValid 置真（合法空工况）；
              ③ 效率按百分数折算，不做效率外推补偿。
*)
FUNCTION FC_DL_ExtrusionBilletHeatCalc : REAL
VAR_INPUT
    fBilletKg  : REAL;   (* 单锭质量 [kg] Billet mass *)
    fCpKJkgK   : REAL;   (* 铝比热容 [kJ/(kg·K)] Aluminium specific heat *)
    fT0C       : REAL;   (* 入炉锭温 [°C] Billet inlet temperature *)
    fT1C       : REAL;   (* 目标出炉锭温 [°C] Billet target temperature *)
    fEffPct    : REAL;   (* 感应加热总效率 [%] Overall induction efficiency *)
    fHeatTimeS : REAL;   (* 允许加热时长 [s] Allowed heating time *)
    nBilletCnt : INT;    (* 同时加热锭数 [件] Number of billets *)
END_VAR
VAR_OUTPUT
    fDeltaTK  : REAL;   (* 单锭温升 [K] Temperature rise per billet *)
    fPowerKW  : REAL;   (* 所需电功率（含效率折算） [kW] Electrical power required *)
    fEnergyKWh: REAL;   (* 本批总电耗 [kWh] Total electrical energy *)
    xValid    : BOOL;   (* 计算有效性标志 [-] Calculation valid flag *)
END_VAR
VAR CONSTANT
    DL_EPS      : REAL := 1.0E-9;   (* 除零判定容差 [无量纲] Divide-by-zero tolerance *)
    DL_KWH_KJ   : REAL := 3600.0;   (* 千焦转千瓦时换算系数 [kJ/kWh] kJ per kWh *)
    DL_PCT_BASE : REAL := 100.0;    (* 百分比基准 [%] Percent base *)
    DL_ZERO     : REAL := 0.0;      (* 零常量 [无量纲] Zero constant *)
END_VAR
VAR
    fHeatKJ  : REAL;   (* 本批所需热量 [kJ] Required heat of the batch *)
    fEffUnit : REAL;   (* 效率折算系数 [-] Efficiency as fraction *)
END_VAR
(* 出口预置：四出口统一预置 *)
fDeltaTK := 0.0; fPowerKW := 0.0; fEnergyKWh := 0.0; xValid := FALSE;
(* 非有限拦截：自反判 NaN，自身差值判 Inf *)
IF (fBilletKg <> fBilletKg) OR ((fBilletKg - fBilletKg) <> 0.0)
   OR (fCpKJkgK <> fCpKJkgK) OR ((fCpKJkgK - fCpKJkgK) <> 0.0)
   OR (fT0C <> fT0C) OR ((fT0C - fT0C) <> 0.0)
   OR (fT1C <> fT1C) OR ((fT1C - fT1C) <> 0.0)
   OR (fEffPct <> fEffPct) OR ((fEffPct - fEffPct) <> 0.0)
   OR (fHeatTimeS <> fHeatTimeS) OR ((fHeatTimeS - fHeatTimeS) <> 0.0) THEN
    FC_DL_ExtrusionBilletHeatCalc := -1.0;  (* 哨兵 -1：输入非有限 / Sentinel -1 non-finite *)
    RETURN;
END_IF
(* 组态域闸：质量/比热/时长/效率/锭数逐引脚覆盖 *)
IF (fBilletKg <= DL_EPS) OR (fCpKJkgK <= DL_EPS) OR (fHeatTimeS <= DL_EPS)
   OR (fEffPct <= DL_ZERO) OR (fEffPct > DL_PCT_BASE) OR (nBilletCnt < 1) THEN
    FC_DL_ExtrusionBilletHeatCalc := -1.0;  (* 哨兵 -1：组态非法 / Sentinel -1 bad config *)
    RETURN;
END_IF
fEffUnit := fEffPct / DL_PCT_BASE;          (* 效率折算为小数 [-] / Efficiency as fraction *)
fDeltaTK := fT1C - fT0C;                    (* 单锭温升 [K] / Temperature rise *)
IF fDeltaTK <= DL_ZERO THEN
    xValid := TRUE;                         (* 合法空工况：无需加热 / Legal no-heating case *)
    FC_DL_ExtrusionBilletHeatCalc := DL_ZERO;
    RETURN;
END_IF
(* 本批热量：Q = n * m * cp * dT [kJ] *)
fHeatKJ := INT_TO_REAL(nBilletCnt) * fBilletKg * fCpKJkgK * fDeltaTK;
(* 电功率：热功率 / 效率，kJ/s = kW *)
fPowerKW := (fHeatKJ / fHeatTimeS) / fEffUnit;
(* 电耗：kJ 除以 3600 得 kWh，效率折算进热量侧 *)
fEnergyKWh := (fHeatKJ / fEffUnit) / DL_KWH_KJ;
xValid := TRUE;                             (* 链路有效 / Chain valid *)
FC_DL_ExtrusionBilletHeatCalc := fPowerKW;  (* 返回电功率 [kW] / Return electrical power *)
END_FUNCTION
